// TIA Portal V18 program export: 5 tag tables, 14 data types, 1 data blocks, 8 code blocks (in call order from the OBs), 0 instance data blocks

VAR_GLOBAL   // PLC tag table "BYPASS_APERTADEIRAS"
   start AT %I1500.1 : Bool;
   remover AT %I1500.2 : Bool;
   reset AT %I1500.3 : Bool;
   MOD1_OK AT %Q1594.0 : Bool;
   MOD2_OK AT %Q1594.1 : Bool;
   RESET_MOD_1 AT %M9.1 : Bool;
   RESET_MOD_2 AT %M9.2 : Bool;
   VALIDACA0_MOD1 AT %M9.6 : Bool;
   VALIDAÇÃO_MOD2 AT %M12.0 : Bool;
   VALIDACAO_ANDON_MOD2 AT %M12.2 : Bool;
   VALIDACAO_ANDON_MOD1 AT %M12.3 : Bool;
   LEANDRO AT %M12.4 : Bool;
   BYPASS_ABST_OLEO AT %M12.6 : Bool;
   BYPASS_ABSTECIMENTO_OLEO AT %M12.7 : Bool;
   BYPASS_ESTANQ_CIL AT %M13.0 : Bool;
   BYPASS_SUP_FREIO AT %M2.1 : Bool;
   BYPASS_PY_EXCENTRICO AT %M2.2 : Bool;
   BYPASS_AP_HARPA AT %M12.5 : Bool;
   BYPASS_BUJAO AT %M13.1 : Bool;
   BYPASS_AP_BUJAO AT %M13.2 : Bool;
   BYPASS_TUBO_RPX AT %M13.3 : Bool;
   BYPASS_AP_TUBO_RPX AT %M13.4 : Bool;
   BYPASS_MOLA_HARPA AT %M13.5 : Bool;
   BYPASS_CARCACA AT %M13.6 : Bool;
   BYPASS_AP_CARCA AT %M13.7 : Bool;
   BYPASS_TALHA_DIF AT %M28.0 : Bool;
   BYPASS_SENSOR_TALHA_DIF AT %M28.1 : Bool;
   BYPASS_PYJUNTA AT %M28.2 : Bool;
   BYPASS_PY_JUNTA AT %M28.3 : Bool;
   BYPASS_CRAWFOOT AT %M28.4 : Bool;
   BYPASS_AP_CRAWFOOT AT %M28.5 : Bool;
   BYPASS_DUPLO_FUSO AT %M28.6 : Bool;
   BYPASS_AP_DUPLO_FUSO AT %M28.7 : Bool;
   BYPASS_P_ESCONDIDA AT %M29.0 : Bool;
   BYPASS_AP_PORCA_ESCON AT %M29.1 : Bool;
   BYPASS_SUP_CIL AT %M29.2 : Bool;
   BYPASS_AP_SUP_CIL AT %M29.3 : Bool;
   BYPASS_PORCA_CIL AT %M29.4 : Bool;
   BYPASS_AP_PORCA_CIL AT %M29.5 : Bool;
   BYPASS_AP_SUP_FREIO AT %M29.6 : Bool;
   BYPASS_PYEXCENTRICO AT %M29.7 : Bool;
   BYPASS_CUBO_DISC AT %M30.0 : Bool;
   BYPASS_PY_CUBO_DISC AT %M30.1 : Bool;
   BYPASS_HOLDER AT %M30.2 : Bool;
   BYPASS_AP_HOLDER AT %M30.3 : Bool;
   BYPASS_CALIPER AT %M30.4 : Bool;
   BYPASS_AP_CALPER AT %M30.5 : Bool;
   BYPASS_PYCUBO_TAMBOR AT %M30.6 : Bool;
   BYPASS_PY_CUBO_TAMBOR AT %M30.7 : Bool;
   BYPASS_HASTE_ALV AT %M31.0 : Bool;
   BYPASS_AP_HASTE_ALV AT %M31.1 : Bool;
   BYPASS_APCUBO AT %M31.2 : Bool;
   BYPASS_AP_CUBO AT %M31.3 : Bool;
   BYPASS_CRAVADOR AT %M31.4 : Bool;
   BYPASS_AP_CRAVADOR AT %M31.5 : Bool;
   BYPASS_INDICADOR AT %M31.6 : Bool;
   BYPASS_AP_INDICADOR AT %M31.7 : Bool;
   BYPASS_VALVULA AT %M32.0 : Bool;
   BYPASS_AP_VALVULA AT %M32.1 : Bool;
   BYPASS_HELGE AT %M32.2 : Bool;
   BYPASS_PY_HELGE AT %M32.3 : Bool;
   BYPASS_PORCA_TERMINAL AT %M32.4 : Bool;
   BYPASS_AP_PORCA_TERMINAL AT %M32.5 : Bool;
   BYPASS_FILTRO_OLEO AT %M32.6 : Bool;
   BYPASS_AP_FILTRO_OLEO AT %M32.7 : Bool;
   BYPASS_REDUCAO AT %M33.0 : Bool;
   BYPASS_AP_REDUCAO AT %M33.1 : Bool;
   BYPASS_FLANGE AT %M33.2 : Bool;
   BYPASS_AP_FLANGE AT %M33.3 : Bool;
   BYPASS_ESTANQ_CILINDRO AT %M33.4 : Bool;
   BYPASS_ESTANQ_CARC AT %M33.5 : Bool;
   BYPASS_ESTANQ_CARCACA AT %M33.6 : Bool;
   EMERG_CABINE_ACIONADA AT %M35.1 : Bool;
   BYPASS_VALVULA_P50 AT %M35.6 : Bool;
   BYPASS_TAMPA_CALIPER_1 AT %M36.0 : Bool;
   BYPASS_AP_VALVULA_P50 AT %M36.1 : Bool;
   TESTE_LEITOR AT %M42.4 : Bool;
   IG_CONTROL_T AT %M43.7 : Bool;
   ABORTA_P05 AT %M2.5 : Bool;
   ABORTA_JOB_P05 AT %M2.6 : Bool;
   TORQUE_ATLAS6000_P15 AT %MD48 : Real;
   PULSO_BORDA_BYPASS AT %M3.1 : Bool;
   BORDA_BYPASS_AP AT %M3.2 : Bool;
   TORQUE_DUPLO_FUSO1 AT %MD52 : Real;
   AUX_APDP AT %M3.4 : Bool;
   SIGNAL_LOST_POKA_JUNTA AT %M3.5 : Bool;
   aux_inicio_receita_pky_p30 AT %M3.7 : Bool;
   JOBOK_POKA_JUNTA_P30 AT %M4.0 : Bool;
   BYPASS_TORQUIMETRO_DIGITAL_1 AT %M4.1 : Bool;
   BYPASS_REULAGEM_ALAVANCA_1 AT %M4.5 : Bool;
   antecipa_expedicao AT %M4.6 : Bool;
   SIGINAL_LOST_PCUBO AT %M5.0 : Bool;
   pulso_teste AT %M5.7 : Bool;
   JOBDONE_ABSTECIMENTO_OLEO AT %M7.3 : Bool;
   SIGNAL_LOST_ABAST_OLEO AT %M7.4 : Bool;
   Bypass_oring_P100 AT %M7.5 : Bool;
   BYPASS_ORING_MAP_P100 AT %M8.1 : Bool;
   SIGNAL_LOST_ORING_MAP AT %M8.3 : Bool;
   InputAuxEdi AT %M8.7 : Bool;
   InputAuxEtr AT %M9.0 : Bool;
   SEM_JOB_PY_OLEO AT %M56.6 : Bool;
   JOB_PY_OLEO AT %M56.7 : Bool;
   JOBDONE_PY_GRAXA AT %M57.2 : Bool;
   Bypass_jidoka_filtro AT %M57.3 : Bool;
   BYPASS_JIDOKA_FILTRO_OLEO_P125 AT %M57.4 : Bool;
   Bypass_vaselina AT %M57.5 : Bool;
   JobOK_vaselina AT %M57.6 : Bool;
   BYpassVaselina AT %M57.7 : Bool;
   resetsinais AT %M58.0 : Bool;
   Bypass_apcilin_pneumatico AT %M58.2 : Bool;
   Bypass_apcilin_pneumaticoP105 AT %M58.3 : Bool;
END_VAR

VAR_GLOBAL   // PLC tag table "BYPASS_STATIONS"
   BYPASS_STATION_1 AT %M36.2 : Bool;
   BYPASS_POSTO_1 AT %M36.3 : Bool;
   BYPASS_STATION_5 AT %M36.4 : Bool;
   BYPASS_POSTO_5 AT %M36.5 : Bool;
   BYPASS_STATION_10 AT %M36.6 : Bool;
   BYPASS_POSTO_10 AT %M36.7 : Bool;
   BYPASS_STATION_15 AT %M37.0 : Bool;
   BYPASS_POSTO_15 AT %M37.1 : Bool;
   BYPASS_STATION_20 AT %M37.2 : Bool;
   BYPASS_POSTO_20 AT %M37.3 : Bool;
   BYPASS_STATION_30 AT %M37.4 : Bool;
   BYPASS_POSTO_30 AT %M37.5 : Bool;
   BYPASS_STATION_40 AT %M37.6 : Bool;
   BYPASS_POSTO_40 AT %M37.7 : Bool;
   BYPASS_STATION_50 AT %M38.0 : Bool;
   BYPASS_POSTO_50 AT %M38.1 : Bool;
   BYPASS_STATION_55 AT %M38.2 : Bool;
   BYPASS_POSTO_55 AT %M38.3 : Bool;
   BYPASS_STATION_60 AT %M38.4 : Bool;
   BYPASS_POSTO_60 AT %M38.5 : Bool;
   BYPASS_STATION_70 AT %M38.6 : Bool;
   BYPASS_POSTO_70 AT %M38.7 : Bool;
   BYPASS_STATION_75 AT %M39.0 : Bool;
   BYPASS_POSTO_75 AT %M39.1 : Bool;
   BYPASS_STATION_80 AT %M39.2 : Bool;
   BYPASS_POSTO_80 AT %M39.3 : Bool;
   BYPASS_STATION_90 AT %M39.4 : Bool;
   BYPASS_POSTO_90 AT %M39.5 : Bool;
   BYPASS_STATION_95 AT %M39.6 : Bool;
   BYPASS_POSTO_95 AT %M39.7 : Bool;
   BYPASS_STATION_100 AT %M40.0 : Bool;
   BYPASS_POSTO_100 AT %M40.1 : Bool;
   BYPASS_STATION_105 AT %M40.2 : Bool;
   BYPASS_POSTO_105 AT %M40.3 : Bool;
   BYPASS_STATION_110 AT %M40.4 : Bool;
   BYPASS_POSTO_110 AT %M40.5 : Bool;
   BYPASS_STATION_115 AT %M40.6 : Bool;
   BYPASS_POSTO_115 AT %M40.7 : Bool;
   BYPASS_STATION_120 AT %M41.0 : Bool;
   BYPASS_POSTO_120 AT %M41.1 : Bool;
   BYPASS_STATION_125 AT %M41.2 : Bool;
   BYPASS_POSTO_125 AT %M41.3 : Bool;
   BYPASS_STATION_130 AT %M41.4 : Bool;
   BYPASS_POSTO_130 AT %M41.5 : Bool;
   BYPASS_STATION_140 AT %M41.6 : Bool;
   BYPASS_POSTO_140 AT %M41.7 : Bool;
   BYPASS_STATION_150 AT %M42.0 : Bool;
   BYPASS_POSTO_150 AT %M42.1 : Bool;
   BYPASS_STATION_QG AT %M42.2 : Bool;
   BYPASS_POSTO_QG AT %M42.3 : Bool;
END_VAR

VAR_GLOBAL   // PLC tag table "Default tag table"
   Forced_WO AT %I1500.0 : Bool;
   Trig_Buffer_ADIC AT %I1500.4 : Bool;
   Trig_Buffer_REMOV AT %I1500.5 : Bool;
   senor_filtro_oleo AT %I1000.0 : Bool;
   LEITOR_LEN AT %IB2283 : Byte;
   LEITURA_DONE AT %I2002.4 : Bool;
   sensor_vaselina AT %I1000.4 : Bool;
   Gatilho_ap_pneumaticaP105 AT %I221.6 : Bool;
   Sensor_RX1_RBX1 AT %I201.7 : Bool;
   Sensor_RX2_RBX2 AT %I201.6 : Bool;
   Sensor_cotovelo_mangueira AT %I1050.0 : Bool;
   Sensor_cotovelo AT %I1050.2 : Bool;
   Sensor_cotovelo_AD1600 AT %I1050.4 : Bool;
   Sensor_plug AT %I1050.6 : Bool;
   Tag_1 AT %QD1302 : DWord;
   Tag_2 AT %Q400.0 : Bool;
   Tag_3 AT %QW1310 : Int;
   SINAL_AP_SEMPRE_LIGADO AT %Q4000.0 : Bool;
   Tag_4 AT %QB1100 : Byte;
   RESET_DESOUTTER_P50 AT %Q8000.0 : Bool;
   RESET_DESOUTTER_P40 AT %Q6000.0 : Bool;
   Limpa_leitor AT %Q2000.7 : Bool;
   Buzzer_P01 AT %Q3.4 : Bool;
   Led_azul_P01 AT %Q3.2 : Bool;
   Led_red_P01 AT %Q3.0 : Bool;
   Led_verde_P01 AT %Q3.1 : Bool;
   Ledverde AT %Q1000.2 : Bool;
   Ledlaranja AT %Q1000.3 : Bool;
   LedVerde_vaselina AT %Q1000.6 : Bool;
   LedAmarelo_vaselina AT %Q1000.7 : Bool;
   LED_RX1_RBX1 AT %Q200.7 : Bool;
   LED_RX2_RBX2 AT %Q200.6 : Bool;
   Buzzer_P40 AT %Q5.4 : Bool;
   Led_azulP40 AT %Q5.2 : Bool;
   Led_VermelhoP40 AT %Q5.0 : Bool;
   Led_VerdeP40 AT %Q5.1 : Bool;
   Led_cotovelo_mangueira AT %Q1050.1 : Bool;
   Led_Cotovelo AT %Q1050.3 : Bool;
   Led_cotovelo_AD1600 AT %Q1050.5 : Bool;
   Led_Plug AT %Q1050.7 : Bool;
   FirstScan AT %M1.0 : Bool;
   DiagStatusUpdate AT %M1.1 : Bool;
   AlwaysTRUE AT %M1.2 : Bool;
   AlwaysFALSE AT %M1.3 : Bool;
   Clock_Byte AT %MB0 : Byte;
   Clock_10Hz AT %M0.0 : Bool;
   Clock_5Hz AT %M0.1 : Bool;
   "Clock_2.5Hz" AT %M0.2 : Bool;
   Clock_2Hz AT %M0.3 : Bool;
   "Clock_1.25Hz" AT %M0.4 : Bool;
   Clock_1Hz AT %M0.5 : Bool;
   "Clock_0.625Hz" AT %M0.6 : Bool;
   "Clock_0.5Hz" AT %M0.7 : Bool;
   status_10 AT %M1.4 : Bool;
   status_20 AT %M1.5 : Bool;
   status_40 AT %M1.6 : Bool;
   status_50 AT %M1.7 : Bool;
   status_60 AT %M6.0 : Bool;
   status_70 AT %M6.1 : Bool;
   status_80 AT %M6.2 : Bool;
   status_90 AT %M6.3 : Bool;
   status_100 AT %M6.4 : Bool;
   status_110 AT %M6.5 : Bool;
   status_120 AT %M6.6 : Bool;
   status_130 AT %M6.7 : Bool;
   BUSY AT %M7.6 : Bool;
   CYCLE_DONE_AREA_IHM AT %M8.0 : Bool;
   MODEZONE_DONE_AREA_IHM AT %M8.2 : Bool;
   CYCLE_DONE_IT_IHM AT %M8.4 : Bool;
   BOTAO_ACIONAR_MENSAGENS AT %M8.5 : Bool;
   Quantity_ok AT %MW10 : Int;
   BYPASSLEITOR AT %M7.7 : Bool;
   Inicia_apertadeiras AT %M4.4 : Bool;
   FORÇA_RECEITA_GERAL AT %M12.1 : Bool;
   CU_PRIMEIRO_POSTO AT %MW14 : Int;
   "POPID_INICO DE_LINHA" AT %M18.0 : LInt;
   Ready_to_copy AT %M2.0 : Bool;
   BYPASS_MOD_2 AT %M2.3 : Bool;
   BYPASS_MOD_1 AT %M2.4 : Bool;
   BYPASS_GERAL_EQUIP AT %M900.1 : Bool;
   "NOVO TESTE" AT %M9.5 : Bool;
   BYPASS_GERAL AT %M33.7 : Bool;
   ESVAZIAMENTO_FALCARE AT %M34.0 : Bool;
   ESVAZIA_FALCARE AT %M34.1 : Bool;
   ESVAZIA_MAIN_LINE AT %M34.2 : Bool;
   ESVAZIAMENTO_MAIN_LINE AT %M34.3 : Bool;
   ESVAZIA_FALCARE_1 AT %M34.4 : Bool;
   ESVAZIA_MAIN_LINE_1 AT %M34.5 : Bool;
   ERRO_ESVAZIAMENTO_LINHA AT %M34.6 : Bool;
   "CABINE EM MANUAL" AT %M34.7 : Bool;
   PRODUCAO_CONCLUIDA AT %M35.0 : Bool;
   GAP_E_EIXO_PENDURADO AT %M35.2 : Bool;
   VALIDACAO_EMERG_MOD1 AT %M35.3 : Bool;
   VALIDACAO_EMERG_MOD2 AT %M35.4 : Bool;
   "SINAL_DE RESET_GAP_CABINE" AT %M35.5 : Bool;
   BYPASS_TAMPA_CALIPER AT %M35.7 : Bool;
   INDEX_LEITOR AT %MW44 : UInt;
   CARACTER AT %MW46 : Int;
   RET_VAL AT %MW200 : Int;
   BYPASS_CABINE_EM_MODO_LOCAL AT %M42.5 : Bool;
   BYPASS_CAB_MODO_LOCAL AT %M42.6 : Bool;
   ACIONA_TELA AT %M43.1 : Bool;
   ERROR_COMUNICACAO_CABINE_SEND AT %M43.2 : Bool;
   ERROR_COMUNICACAO_CABINE_RECIVE AT %M43.3 : Bool;
   BYPASS_LEITURA AT %M43.4 : Bool;
   BORDA_MODZ1 AT %M43.5 : Bool;
   BYPASS_PY_JUNTA_RX_RBX AT %M43.6 : Bool;
   bypass_sem_receita AT %M2.7 : Bool;
   provisorio AT %M3.0 : Bool;
   BYPASS_PRENSA_LEMARB AT %M3.3 : Bool;
   TOOLRUNNING_POKA_JUNTA AT %M3.6 : Bool;
   BYPASS_TORQUIMETRO_DIGITAL AT %M4.2 : Bool;
   BYPASS_REULAGEM_ALAVANCA AT %M4.3 : Bool;
   ATIVA_FOR AT %M4.7 : Bool;
   PULSO_BY_P110 AT %M5.1 : Bool;
   set_modezone_done AT %M5.2 : Bool;
   giro_cabine AT %M5.3 : Bool;
   cabine_rodou AT %M5.4 : Bool;
   reset_md1 AT %M5.5 : Bool;
   reset_md2 AT %M5.6 : Bool;
   aux_gap AT %M7.0 : Bool;
   guarda_gap AT %M7.1 : Bool;
   chamada_forcada AT %MW16 : Int;
   Cabin_line_reference AT %M7.2 : Bool;
   SIGNAL_LOST_HELGE_2 AT %M8.6 : Bool;
   Habilita_matrix_P01 AT %M9.3 : Bool;
   Habilita_matrix_P05 AT %M9.4 : Bool;
   Habilita_matrix_P10 AT %M9.7 : Bool;
   Habilita_matrix_P15 AT %M26.0 : Bool;
   Habilita_matrix_P20 AT %M26.1 : Bool;
   Habilita_matrix_P30 AT %M26.2 : Bool;
   Habilita_matrix_P40 AT %M26.3 : Bool;
   Habilita_matrix_P50 AT %M26.4 : Bool;
   Habilita_matrix_P55 AT %M26.5 : Bool;
   Habilita_matrix_P60 AT %M26.6 : Bool;
   Habilita_matrix_P70 AT %M26.7 : Bool;
   Habilita_matrix_P75 AT %M27.0 : Bool;
   Habilita_matrix_P80 AT %M27.1 : Bool;
   Habilita_matrix_P90 AT %M27.2 : Bool;
   Habilita_matrix_P95 AT %M27.3 : Bool;
   Habilita_matrix_P100 AT %M27.4 : Bool;
   Habilita_matrix_P105 AT %M27.5 : Bool;
   Habilita_matrix_P110 AT %M27.6 : Bool;
   Habilita_matrix_P115 AT %M27.7 : Bool;
   Habilita_matrix_P120 AT %M42.7 : Bool;
   Habilita_matrix_P125 AT %M43.0 : Bool;
   Habilita_matrix_P130 AT %M56.0 : Bool;
   Habilita_matrix_P140 AT %M56.1 : Bool;
   Habilita_matrix_P150 AT %M56.2 : Bool;
   Habilita_matrix_QG AT %M56.3 : Bool;
   Bypass_graxa AT %M56.4 : Bool;
   Bypass_graxa_expedicao AT %M56.5 : Bool;
   JOBOK_PY_OLEO AT %M57.0 : Bool;
   antecipa_expedicao_1 AT %M57.1 : Bool;
   bahia AT %M58.1 : Bool;
   Count_gatilho AT %MW60 : Int;
END_VAR
VAR_GLOBAL CONSTANT   // user constants
   Config_OPC : Int := 17;
   maxConnectionsOPCUA : Int := 5;
END_VAR

VAR_GLOBAL   // PLC tag table "LEITOR_VIVERK"
   Readcomplete AT %I2000.1 : Bool;
   ResultData0 AT %IB2284 : Byte;
   ResultData1 AT %IB2285 : Byte;
   ResultData2 AT %IB2286 : Byte;
   ResultData3 AT %IB2287 : Byte;
   ResultData4 AT %IB2288 : Byte;
   ResultData5 AT %IB2289 : Byte;
   ResultData6 AT %IB2290 : Byte;
   ResultData7 AT %IB2291 : Byte;
   ResultData8 AT %IB2292 : Byte;
   ResultData9 AT %IB2293 : Byte;
   ResultData10 AT %IB2294 : Byte;
   ResultData11 AT %IB2295 : Byte;
   ResultData12 AT %IB2296 : Byte;
   Tag_5 AT %IB2000 : Byte;
   Tag_6 AT %IB2001 : Byte;
   Tag_7 AT %IB2002 : Byte;
   Tag_8 AT %IB2003 : Byte;
   Tag_9 AT %IB2004 : Byte;
   Tag_10 AT %IB2005 : Byte;
   Tag_11 AT %IB2006 : Byte;
   Tag_12 AT %IB2007 : Byte;
   Tag_13 AT %IB2008 : Byte;
   Tag_14 AT %IB2009 : Byte;
   Tag_15 AT %IB2010 : Byte;
   Tag_16 AT %IB2011 : Byte;
   Tag_17 AT %IB2012 : Byte;
   Tag_18 AT %IB2013 : Byte;
END_VAR

VAR_GLOBAL   // PLC tag table "Setup"
   Tag_19 AT %I0.0 : Bool;
END_VAR
VAR_GLOBAL CONSTANT   // user constants
   ModeZone_Setup_Const : Int := 12;
   Station_Setup_Const : Int := 20;
   Position_Setup_Const : Int := 1;
   Equipment_Setup_Const : Int := 10;
   ThisProcess : Int := 1;
   ThisWorkshop : Int := 1;
   Connection_Setup_Const : Int := 30;
   ContractID_Setup_Const : Int := 24;
   ITConnectionName : String := 'PLC_AREA_01';
   Parameter_Setup_Const : Int := 20;
   WorkPlace_Setup_Const : Int := 16;
   Total_User_Const : Int := 200;
   User_Roles_Const : Int := 100;
   ProductionSequenceList_Setup_Const : Int := 30;   // Quantidade de produtos que podemos ter por posto
   listTypeReason_Const : Int := 200;
   ITConnectionID : Word := W#16#101;
   Signal_Setup_Const : Int := 8;
   ShiftList_Setup_Const : Int := 3;
   Quantidade_task : Int := 10;
   Tamanho_POPID : Int := 7;
   nProcess : Int := 1;
   Quantidade_Paradas_Matriz : Int := 2;
END_VAR

TYPE "Comm"
   STRUCT
      Connection_ID : Word;
      R_ID : CONN_R_ID;
      REQ : Bool;
      Len : Word;
      Result : Struct
         DONE : Bool;
         ERROR : Bool;
         STATUS : Word;
      END_STRUCT;
      Diagnostic : Struct
         countDone : Int;
         countError : Int;
         memStatus : Word;
      END_STRUCT;
   END_STRUCT;
END_TYPE

TYPE "Config_SEND_RCV"
   STRUCT
      modezone { S7_SetPoint := 'True'} : Array[1.."ModeZone_Setup_Const"] of "Comm";
   END_STRUCT;
END_TYPE

TYPE "InterlockEmergMdz_in"
   STRUCT
      StationInterlock_APLC_Input : Array[1.."Station_Setup_Const"] of Struct
         Emergencial_Interlock_APLC_Input : Bool;
      END_STRUCT;
   END_STRUCT;
END_TYPE

TYPE "InterlockMdz_in"
   STRUCT
      StationInterlock_APLC_Input : Array[1.."Station_Setup_Const"] of Struct
         PositionInterlock_APLC_Input : Array[1.."Position_Setup_Const"] of Struct
            LoginInterlock_APLC : Bool;
            EquipmentInterlock_APLC_Input : Array[1.."Equipment_Setup_Const"] of Struct
               SignalInterlock_APLC_Input : Array[1.."Signal_Setup_Const"] of Bool;
            END_STRUCT;
         END_STRUCT;
      END_STRUCT;
   END_STRUCT;
END_TYPE

TYPE "Modezone_Gap"
   STRUCT
      GapActive : Bool;
   END_STRUCT;
END_TYPE

TYPE "Process_Gap"
   STRUCT
      ProcessGapActive : Bool;
      ModezoneGap { S7_SetPoint := 'True'} : Array[1.."ModeZone_Setup_Const"] of "Modezone_Gap";
   END_STRUCT;
END_TYPE

TYPE "TaktModeZone_Input"
   STRUCT
      ModeZone_Done : Bool;
   END_STRUCT;
END_TYPE

TYPE "TargetProductionMdz_in"
   STRUCT
      KPI_Informations : Struct
         Full_AvailabilityShift : Array[1.."ShiftList_Setup_Const"] of Time;
         Full_AvailabilityDay : Time := T#9H_15M;
         Net_AvailabilityShift : Array[1.."ShiftList_Setup_Const"] of Time;
         Net_AvailabilityDay : Time := T#9H_15M;
         Total_StopPlannedShift : Array[1.."ShiftList_Setup_Const"] of Time;
         Total_StopPlannedDay : Time := T#0MS;
         StopPlanned_Executed_Shift : Array[1.."ShiftList_Setup_Const"] of Time;
         StopPlanned_Executed_Day : Time := T#2H_45M;
         NextStopPlanned : Date_And_Time := DT#2000-01-10-00:00:00;
         NextStopPlanned_Index : Int := 11;
         RemaningTimeToStopPlanned : Time := T#8D_15H_45M_48S_109MS;
         NextStopPlannedInRealTime : Time := T#8H_14M_11S_891MS;
         RemaningCycleToStoPplanned : DInt := 2_139_095_040;
         Total_StopTimeShift : Array[1.."ShiftList_Setup_Const"] of Time;
         Total_StopTimeDay : Time := T#-1H_41M_28S;
         GoalOfShift : Array[1.."ShiftList_Setup_Const"] of Int;
         GoalOfDay : Int := 199;
         TaktStandardByShift : Array[1.."ShiftList_Setup_Const"] of Time;
      END_STRUCT;
      KPI_Results : Struct
         Production_Status : Int := 0;
         MaxProductionCapacity_Shift : Array[1.."ShiftList_Setup_Const"] of Int;
         MaxProductionCapacity_Day : Int := 246;
         TimeToProductionDone_Shift : Array[1.."ShiftList_Setup_Const"] of Time;
         TimeToProductionDone_Day : Time := T#0MS;
      END_STRUCT;
   END_STRUCT;
   // KPI_Informations.Full_AvailabilityShift[1] := T#9H_15M;
   // KPI_Informations.Full_AvailabilityShift[2..3] := T#0MS;
   // KPI_Informations.Net_AvailabilityShift[1] := T#9H_15M;
   // KPI_Informations.Net_AvailabilityShift[2..3] := T#0MS;
   // KPI_Informations.Total_StopPlannedShift[1..3] := T#0MS;
   // KPI_Informations.StopPlanned_Executed_Shift[1] := T#1H_35M;
   // KPI_Informations.StopPlanned_Executed_Shift[2] := T#1H_10M;
   // KPI_Informations.StopPlanned_Executed_Shift[3] := T#0MS;
   // KPI_Informations.Total_StopTimeShift[1] := T#-1H_11M_58S;
   // KPI_Informations.Total_StopTimeShift[2] := T#-29M_30S;
   // KPI_Informations.Total_StopTimeShift[3] := T#0MS;
   // KPI_Informations.GoalOfShift[1] := 164;
   // KPI_Informations.GoalOfShift[2] := 35;
   // KPI_Informations.GoalOfShift[3] := 0;
   // KPI_Informations.TaktStandardByShift[1] := T#2M_15S;
   // KPI_Informations.TaktStandardByShift[2] := T#10M;
   // KPI_Informations.TaktStandardByShift[3] := T#0MS;
   // KPI_Results.MaxProductionCapacity_Shift[1] := 246;
   // KPI_Results.MaxProductionCapacity_Shift[2..3] := 0;
   // KPI_Results.TimeToProductionDone_Shift[1..3] := T#0MS;
END_TYPE

TYPE "UDT_DadosEquipScala"
   STRUCT
      Bool0 : Bool;
      Bool1 : Bool;
      Bool2 : Bool;
      Bool3 : Bool;
      Bool4 : Bool;
      Bool5 : Bool;
      Bool6 : Bool;
      Bool7 : Bool;
      Bool8 : Bool;
      Bool9 : Bool;
      Bool10 : Bool;
      Bool11 : Bool;
      Bool12 : Bool;
      Bool13 : Bool;
      Bool14 : Bool;
      Bool15 : Bool;
   END_STRUCT;
END_TYPE

TYPE "UDT_EquipamentoScala"
   STRUCT
      Equipamento : Array[1..18] of "UDT_DadosEquipScala";
   END_STRUCT;
END_TYPE

TYPE "Udt_DataAGVStation"
   STRUCT
      Station { S7_SetPoint := 'True'} : Array[1..20] of "Udt_Data_AGVToScala";
   END_STRUCT;
END_TYPE

TYPE "Udt_Data_AGVToScala"
   STRUCT
      POPID : String[10];   // POPID
      CU : String[10];   // CU
      AGVNumber : Int;   // Número AGV
      ProductOK : Bool;   // Produto recebido OK
      ProductNOK : Bool;   // Falha produto recebido Scala
      AGVRedCard : Bool;   // AGV com trabalho
      Spare4 : Bool;   // Reserva
      Spare5 : Bool;   // Reserva
      Spare6 : Bool;   // Reserva
      Spare7 : Bool;   // Reserva
      Spare8 : Bool;   // Reserva
      Spare9 : Bool;   // Reserva
      Spare10 : Bool;   // Reserva
      Spare11 : Bool;   // Reserva
      Spare12 : Bool;   // Reserva
      Spare13 : Bool;   // Reserva
      Spare14 : Bool;   // Reserva
      Spare15 : Bool;   // Reserva
      Spare16 : Bool;   // Reserva
   END_STRUCT;
END_TYPE

TYPE "UserValidationMdz_in"
   STRUCT
      Station : Array[1.."Station_Setup_Const"] of Struct
         UserMaster_ID : DInt;
         Position_ID_Validation : Int;
         LogIn : Bool;
         Position : Array[1.."Position_Setup_Const"] of Struct
            User_ID : DInt;
            BadgeNumber : LInt;
            LogIn : Bool;
            LogOut : Bool;
            ByPass : Bool;
         END_STRUCT;
      END_STRUCT;
   END_STRUCT;
   // Station[1..20].UserMaster_ID := 0;
   // Station[1..20].Position_ID_Validation := 0;
   // Station[1..20].LogIn := FALSE;
   // Station[1].Position[1].User_ID := 0;
   // Station[2].Position[1].User_ID := 0;
   // Station[3].Position[1].User_ID := 0;
   // Station[4].Position[1].User_ID := 0;
   // Station[5].Position[1].User_ID := 0;
   // Station[6].Position[1].User_ID := 0;
   // Station[7].Position[1].User_ID := 0;
   // Station[8].Position[1].User_ID := 0;
   // Station[9].Position[1].User_ID := 0;
   // Station[10].Position[1].User_ID := 0;
   // Station[11].Position[1].User_ID := 0;
   // Station[12].Position[1].User_ID := 0;
   // Station[13].Position[1].User_ID := 0;
   // Station[14].Position[1].User_ID := 0;
   // Station[15].Position[1].User_ID := 0;
   // Station[16].Position[1].User_ID := 0;
   // Station[17].Position[1].User_ID := 0;
   // Station[18].Position[1].User_ID := 0;
   // Station[19].Position[1].User_ID := 0;
   // Station[20].Position[1].User_ID := 0;
   // Station[1].Position[1].BadgeNumber := 0;
   // Station[2].Position[1].BadgeNumber := 0;
   // Station[3].Position[1].BadgeNumber := 0;
   // Station[4].Position[1].BadgeNumber := 0;
   // Station[5].Position[1].BadgeNumber := 0;
   // Station[6].Position[1].BadgeNumber := 0;
   // Station[7].Position[1].BadgeNumber := 0;
   // Station[8].Position[1].BadgeNumber := 0;
   // Station[9].Position[1].BadgeNumber := 0;
   // Station[10].Position[1].BadgeNumber := 0;
   // Station[11].Position[1].BadgeNumber := 0;
   // Station[12].Position[1].BadgeNumber := 0;
   // Station[13].Position[1].BadgeNumber := 0;
   // Station[14].Position[1].BadgeNumber := 0;
   // Station[15].Position[1].BadgeNumber := 0;
   // Station[16].Position[1].BadgeNumber := 0;
   // Station[17].Position[1].BadgeNumber := 0;
   // Station[18].Position[1].BadgeNumber := 0;
   // Station[19].Position[1].BadgeNumber := 0;
   // Station[20].Position[1].BadgeNumber := 0;
   // Station[1].Position[1].LogIn := FALSE;
   // Station[2].Position[1].LogIn := FALSE;
   // Station[3].Position[1].LogIn := FALSE;
   // Station[4].Position[1].LogIn := FALSE;
   // Station[5].Position[1].LogIn := FALSE;
   // Station[6].Position[1].LogIn := FALSE;
   // Station[7].Position[1].LogIn := FALSE;
   // Station[8].Position[1].LogIn := FALSE;
   // Station[9].Position[1].LogIn := FALSE;
   // Station[10].Position[1].LogIn := FALSE;
   // Station[11].Position[1].LogIn := FALSE;
   // Station[12].Position[1].LogIn := FALSE;
   // Station[13].Position[1].LogIn := FALSE;
   // Station[14].Position[1].LogIn := FALSE;
   // Station[15].Position[1].LogIn := FALSE;
   // Station[16].Position[1].LogIn := FALSE;
   // Station[17].Position[1].LogIn := FALSE;
   // Station[18].Position[1].LogIn := FALSE;
   // Station[19].Position[1].LogIn := FALSE;
   // Station[20].Position[1].LogIn := FALSE;
   // Station[1].Position[1].LogOut := TRUE;
   // Station[2].Position[1].LogOut := TRUE;
   // Station[3].Position[1].LogOut := TRUE;
   // Station[4].Position[1].LogOut := TRUE;
   // Station[5].Position[1].LogOut := TRUE;
   // Station[6].Position[1].LogOut := TRUE;
   // Station[7].Position[1].LogOut := TRUE;
   // Station[8].Position[1].LogOut := TRUE;
   // Station[9].Position[1].LogOut := TRUE;
   // Station[10].Position[1].LogOut := TRUE;
   // Station[11].Position[1].LogOut := TRUE;
   // Station[12].Position[1].LogOut := TRUE;
   // Station[13].Position[1].LogOut := TRUE;
   // Station[14].Position[1].LogOut := TRUE;
   // Station[15].Position[1].LogOut := TRUE;
   // Station[16].Position[1].LogOut := TRUE;
   // Station[17].Position[1].LogOut := TRUE;
   // Station[18].Position[1].LogOut := TRUE;
   // Station[19].Position[1].LogOut := TRUE;
   // Station[20].Position[1].LogOut := TRUE;
   // Station[1].Position[1].ByPass := FALSE;
   // Station[2].Position[1].ByPass := FALSE;
   // Station[3].Position[1].ByPass := FALSE;
   // Station[4].Position[1].ByPass := FALSE;
   // Station[5].Position[1].ByPass := FALSE;
   // Station[6].Position[1].ByPass := FALSE;
   // Station[7].Position[1].ByPass := FALSE;
   // Station[8].Position[1].ByPass := FALSE;
   // Station[9].Position[1].ByPass := FALSE;
   // Station[10].Position[1].ByPass := FALSE;
   // Station[11].Position[1].ByPass := FALSE;
   // Station[12].Position[1].ByPass := FALSE;
   // Station[13].Position[1].ByPass := FALSE;
   // Station[14].Position[1].ByPass := FALSE;
   // Station[15].Position[1].ByPass := FALSE;
   // Station[16].Position[1].ByPass := FALSE;
   // Station[17].Position[1].ByPass := FALSE;
   // Station[18].Position[1].ByPass := FALSE;
   // Station[19].Position[1].ByPass := FALSE;
   // Station[20].Position[1].ByPass := FALSE;
END_TYPE

TYPE "UserValidationMdz_out"
   STRUCT
      Station : Array[1.."Station_Setup_Const"] of Struct
         Position : Array[1.."Position_Setup_Const"] of Struct
            User_ID : DInt;
            User_SSB : String[8];
            UserName : String[37];
            MsgLogin : String[40];
            AuthorizedByUserMaster_ID : DInt;
            Authentication : Bool;
         END_STRUCT;
      END_STRUCT;
   END_STRUCT;
   // Station[1].Position[1].User_ID := 0;
   // Station[2].Position[1].User_ID := 0;
   // Station[3].Position[1].User_ID := 0;
   // Station[4].Position[1].User_ID := 0;
   // Station[5].Position[1].User_ID := 0;
   // Station[6].Position[1].User_ID := 0;
   // Station[7].Position[1].User_ID := 0;
   // Station[8].Position[1].User_ID := 0;
   // Station[9].Position[1].User_ID := 0;
   // Station[10].Position[1].User_ID := 0;
   // Station[11].Position[1].User_ID := 0;
   // Station[12].Position[1].User_ID := 0;
   // Station[13].Position[1].User_ID := 0;
   // Station[14].Position[1].User_ID := 0;
   // Station[15].Position[1].User_ID := 0;
   // Station[16].Position[1].User_ID := 0;
   // Station[17].Position[1].User_ID := 0;
   // Station[18].Position[1].User_ID := 0;
   // Station[19].Position[1].User_ID := 0;
   // Station[20].Position[1].User_ID := 0;
   // Station[1].Position[1].User_SSB := '';
   // Station[2].Position[1].User_SSB := '';
   // Station[3].Position[1].User_SSB := '';
   // Station[4].Position[1].User_SSB := '';
   // Station[5].Position[1].User_SSB := '';
   // Station[6].Position[1].User_SSB := '';
   // Station[7].Position[1].User_SSB := '';
   // Station[8].Position[1].User_SSB := '';
   // Station[9].Position[1].User_SSB := '';
   // Station[10].Position[1].User_SSB := '';
   // Station[11].Position[1].User_SSB := '';
   // Station[12].Position[1].User_SSB := '';
   // Station[13].Position[1].User_SSB := '';
   // Station[14].Position[1].User_SSB := '';
   // Station[15].Position[1].User_SSB := '';
   // Station[16].Position[1].User_SSB := '';
   // Station[17].Position[1].User_SSB := '';
   // Station[18].Position[1].User_SSB := '';
   // Station[19].Position[1].User_SSB := '';
   // Station[20].Position[1].User_SSB := '';
   // Station[1].Position[1].UserName := '';
   // Station[2].Position[1].UserName := '';
   // Station[3].Position[1].UserName := '';
   // Station[4].Position[1].UserName := '';
   // Station[5].Position[1].UserName := '';
   // Station[6].Position[1].UserName := '';
   // Station[7].Position[1].UserName := '';
   // Station[8].Position[1].UserName := '';
   // Station[9].Position[1].UserName := '';
   // Station[10].Position[1].UserName := '';
   // Station[11].Position[1].UserName := '';
   // Station[12].Position[1].UserName := '';
   // Station[13].Position[1].UserName := '';
   // Station[14].Position[1].UserName := '';
   // Station[15].Position[1].UserName := '';
   // Station[16].Position[1].UserName := '';
   // Station[17].Position[1].UserName := '';
   // Station[18].Position[1].UserName := '';
   // Station[19].Position[1].UserName := '';
   // Station[20].Position[1].UserName := '';
   // Station[1].Position[1].MsgLogin := 'POSTO: 1 NAO POSSUI USUARIO CADASTRADO';
   // Station[2].Position[1].MsgLogin := 'POSTO: 1 NAO POSSUI USUARIO CADASTRADO';
   // Station[3].Position[1].MsgLogin := 'POSTO: 1 NAO POSSUI USUARIO CADASTRADO';
   // Station[4].Position[1].MsgLogin := 'POSTO: 1 NAO POSSUI USUARIO CADASTRADO';
   // Station[5].Position[1].MsgLogin := 'POSTO: 1 NAO POSSUI USUARIO CADASTRADO';
   // Station[6].Position[1].MsgLogin := 'POSTO: 1 NAO POSSUI USUARIO CADASTRADO';
   // Station[7].Position[1].MsgLogin := 'POSTO: 1 NAO POSSUI USUARIO CADASTRADO';
   // Station[8].Position[1].MsgLogin := 'POSTO: 1 NAO POSSUI USUARIO CADASTRADO';
   // Station[9].Position[1].MsgLogin := 'POSTO: 1 NAO POSSUI USUARIO CADASTRADO';
   // Station[10].Position[1].MsgLogin := 'POSTO: 1 NAO POSSUI USUARIO CADASTRADO';
   // Station[11].Position[1].MsgLogin := 'POSTO: 1 NAO POSSUI USUARIO CADASTRADO';
   // Station[12].Position[1].MsgLogin := 'POSTO: 1 NAO POSSUI USUARIO CADASTRADO';
   // Station[13].Position[1].MsgLogin := 'POSTO: 1 NAO POSSUI USUARIO CADASTRADO';
   // Station[14].Position[1].MsgLogin := 'POSTO: 1 NAO POSSUI USUARIO CADASTRADO';
   // Station[15].Position[1].MsgLogin := 'POSTO: 1 NAO POSSUI USUARIO CADASTRADO';
   // Station[16].Position[1].MsgLogin := 'POSTO: 1 NAO POSSUI USUARIO CADASTRADO';
   // Station[17].Position[1].MsgLogin := 'POSTO: 1 NAO POSSUI USUARIO CADASTRADO';
   // Station[18].Position[1].MsgLogin := 'POSTO: 1 NAO POSSUI USUARIO CADASTRADO';
   // Station[19].Position[1].MsgLogin := 'POSTO: 1 NAO POSSUI USUARIO CADASTRADO';
   // Station[20].Position[1].MsgLogin := 'POSTO: 1 NAO POSSUI USUARIO CADASTRADO';
   // Station[1].Position[1].AuthorizedByUserMaster_ID := 0;
   // Station[2].Position[1].AuthorizedByUserMaster_ID := 0;
   // Station[3].Position[1].AuthorizedByUserMaster_ID := 0;
   // Station[4].Position[1].AuthorizedByUserMaster_ID := 0;
   // Station[5].Position[1].AuthorizedByUserMaster_ID := 0;
   // Station[6].Position[1].AuthorizedByUserMaster_ID := 0;
   // Station[7].Position[1].AuthorizedByUserMaster_ID := 0;
   // Station[8].Position[1].AuthorizedByUserMaster_ID := 0;
   // Station[9].Position[1].AuthorizedByUserMaster_ID := 0;
   // Station[10].Position[1].AuthorizedByUserMaster_ID := 0;
   // Station[11].Position[1].AuthorizedByUserMaster_ID := 0;
   // Station[12].Position[1].AuthorizedByUserMaster_ID := 0;
   // Station[13].Position[1].AuthorizedByUserMaster_ID := 0;
   // Station[14].Position[1].AuthorizedByUserMaster_ID := 0;
   // Station[15].Position[1].AuthorizedByUserMaster_ID := 0;
   // Station[16].Position[1].AuthorizedByUserMaster_ID := 0;
   // Station[17].Position[1].AuthorizedByUserMaster_ID := 0;
   // Station[18].Position[1].AuthorizedByUserMaster_ID := 0;
   // Station[19].Position[1].AuthorizedByUserMaster_ID := 0;
   // Station[20].Position[1].AuthorizedByUserMaster_ID := 0;
   // Station[1].Position[1].Authentication := FALSE;
   // Station[2].Position[1].Authentication := FALSE;
   // Station[3].Position[1].Authentication := FALSE;
   // Station[4].Position[1].Authentication := FALSE;
   // Station[5].Position[1].Authentication := FALSE;
   // Station[6].Position[1].Authentication := FALSE;
   // Station[7].Position[1].Authentication := FALSE;
   // Station[8].Position[1].Authentication := FALSE;
   // Station[9].Position[1].Authentication := FALSE;
   // Station[10].Position[1].Authentication := FALSE;
   // Station[11].Position[1].Authentication := FALSE;
   // Station[12].Position[1].Authentication := FALSE;
   // Station[13].Position[1].Authentication := FALSE;
   // Station[14].Position[1].Authentication := FALSE;
   // Station[15].Position[1].Authentication := FALSE;
   // Station[16].Position[1].Authentication := FALSE;
   // Station[17].Position[1].Authentication := FALSE;
   // Station[18].Position[1].Authentication := FALSE;
   // Station[19].Position[1].Authentication := FALSE;
   // Station[20].Position[1].Authentication := FALSE;
END_TYPE

DATA_BLOCK "VERIFICA INTERLOCK"   // DB200
{ S7_Optimized_Access := 'TRUE' }
// stored: MemoryReserve 100
   VAR
      INTERLOCK : Array[0..10] of Struct
         STATION : Int;
         EQUIPAMENTO : Int;
         SINAL : Int;
      END_STRUCT;
      "ATIVA FOR" : Bool;
      modezone : Int;
   END_VAR
BEGIN
END_DATA_BLOCK

ORGANIZATION_BLOCK "OB1 Main"   // OB1, LAD, ProgramCycle
TITLE = "Main Program Sweep (Cycle)"
{ S7_Optimized_Access := 'TRUE' }
// stored: SetENOAutomatically false
   VAR_INPUT
      Initial_Call : Bool;   // Initial call of this OB
      Remanence : Bool;   // =True, if remanent data are available
   END_VAR
   VAR_TEMP
      ADR : UDInt;
      LEN : UInt;
      "RETURN" : Int;
      ERROR : Bool;
      STATUS : Word;
      DONE : Bool;
      POPID : String;
      CU : Int;
      Quantidade_erro : Int;
      DONE_MAIN_LINE_PUT : Bool;
      ERROR_MAIN_LINE_PUT : Bool;
      DONE_MAIN_LINE_GET : Bool;
      ERROR_MAIN_LINE_GET : Bool;
      DONE_FALCARE_PUT : Bool;
      ERROR_FALCARE_PUT : Bool;
      DONE_FALCARE_GET : Bool;
      ERROR_FALCARE_GET : Bool;
      DONE_GIRADOR_PUT : Bool;
      ERROR_GIRADOR_PUT : Bool;
      DONE_GIRADOR_GET : Bool;
      ERROR_GIRADOR_GET : Bool;
      DONE_ABSTECIMENTO_OLEO_PUT : Bool;
      ERRO_ABASTECIMENTO_OLEO_PUT : Bool;
      DONE_ABSTECIMENTO_OLEO_GET : Bool;
      ERRO_ABSTECIMENTO_OLEO_GET : Bool;
      ERROR_ALARMS_IHM_FALCARE_GET : Bool;
      DONE_ALARMS_IHM_FALCARE_GET : Bool;
      AUX_BSEND_LEMARB : Word;
      AUX_RECIVE_LEMARB : Word;
   END_VAR
BEGIN

REGION Network 1: Set Id Connection automatic
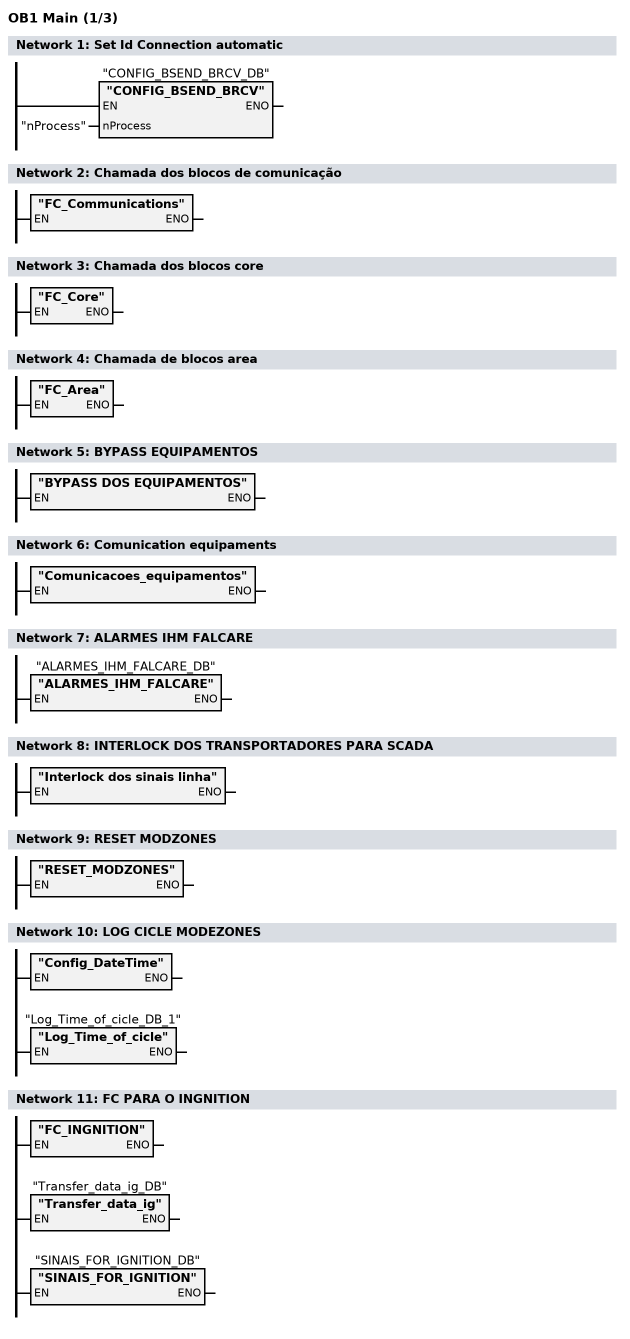
   RUNG wire#powerrail
      "CONFIG_BSEND_BRCV_DB"(nProcess := "nProcess")
   END_RUNG
   // the same network as SCL:
   "CONFIG_BSEND_BRCV_DB"(nProcess := "nProcess");   // "CONFIG_BSEND_BRCV"
END_REGION

REGION Network 2: Chamada dos blocos de comunicação
   RUNG wire#powerrail
      "FC_Communications"()
   END_RUNG
   // the same network as SCL:
   "FC_Communications"();
END_REGION

REGION Network 3: Chamada dos blocos core
   RUNG wire#powerrail
      "FC_Core"()
   END_RUNG
   // the same network as SCL:
   "FC_Core"();
END_REGION

REGION Network 4: Chamada de blocos area
   RUNG wire#powerrail
      "FC_Area"()
   END_RUNG
   // the same network as SCL:
   "FC_Area"();
END_REGION

REGION Network 5: BYPASS EQUIPAMENTOS
   RUNG wire#powerrail
      "BYPASS DOS EQUIPAMENTOS"()
   END_RUNG
   // the same network as SCL:
   "BYPASS DOS EQUIPAMENTOS"();
END_REGION

REGION Network 6: Comunication equipaments
   RUNG wire#powerrail
      "Comunicacoes_equipamentos"()
   END_RUNG
   // the same network as SCL:
   "Comunicacoes_equipamentos"();
END_REGION

REGION Network 7: ALARMES IHM FALCARE
   RUNG wire#powerrail
      "ALARMES_IHM_FALCARE_DB"()
   END_RUNG
   // the same network as SCL:
   "ALARMES_IHM_FALCARE_DB"();   // "ALARMES_IHM_FALCARE"
END_REGION

REGION Network 8: INTERLOCK DOS TRANSPORTADORES PARA SCADA
   RUNG wire#powerrail
      "Interlock dos sinais linha"()
   END_RUNG
   // the same network as SCL:
   "Interlock dos sinais linha"();
END_REGION

REGION Network 9: RESET MODZONES
   RUNG wire#powerrail
      "RESET_MODZONES"()
   END_RUNG
   // the same network as SCL:
   "RESET_MODZONES"();
END_REGION

REGION Network 10: LOG CICLE MODEZONES
   RUNG wire#powerrail
      "Config_DateTime"()
   END_RUNG
   RUNG wire#powerrail
      "Log_Time_of_cicle_DB_1"()
   END_RUNG
   // the same network as SCL:
   "Config_DateTime"();
   "Log_Time_of_cicle_DB_1"();   // "Log_Time_of_cicle"
END_REGION

REGION Network 11: FC PARA O INGNITION
   RUNG wire#powerrail
      "FC_INGNITION"()
   END_RUNG
   RUNG wire#powerrail
      "Transfer_data_ig_DB"()
   END_RUNG
   RUNG wire#powerrail
      "SINAIS_FOR_IGNITION_DB"()
   END_RUNG
   // the same network as SCL:
   "FC_INGNITION"();
   "Transfer_data_ig_DB"();   // "Transfer_data_ig"
   "SINAIS_FOR_IGNITION_DB"();   // "SINAIS_FOR_IGNITION"
END_REGION

REGION Network 12: TESTE DE VALIDAÇÃO MODEZONES
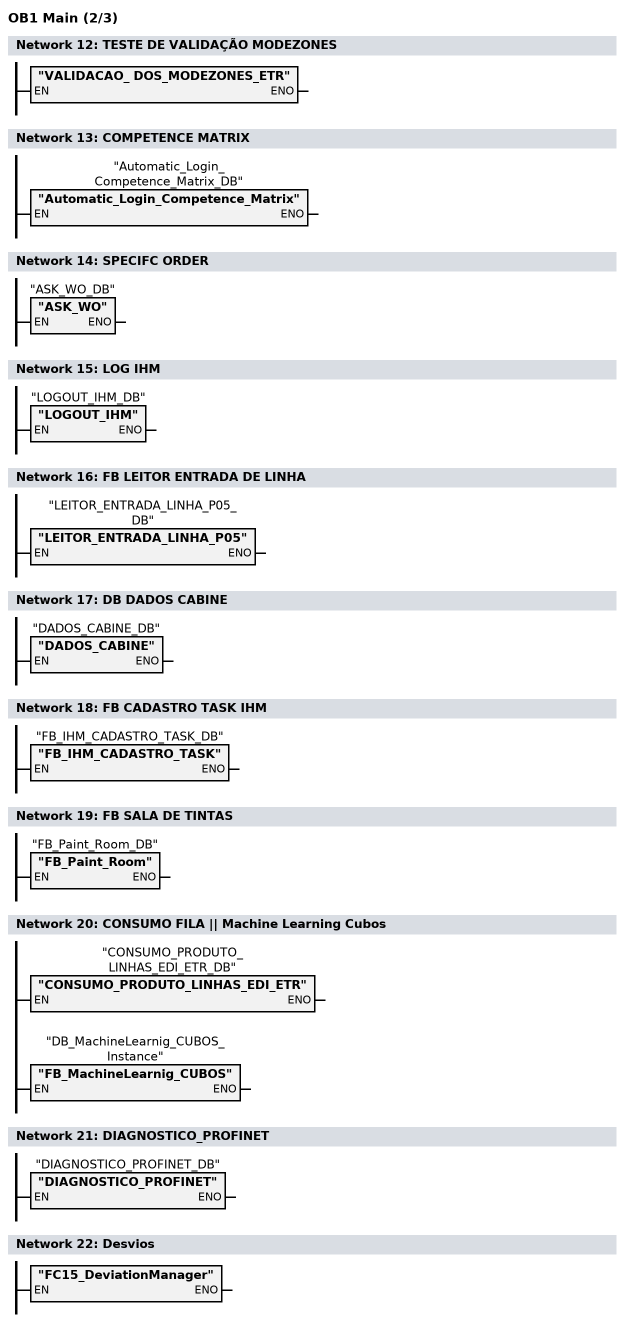
   RUNG wire#powerrail
      "VALIDACAO_ DOS_MODEZONES_ETR"()
   END_RUNG
   // the same network as SCL:
   "VALIDACAO_ DOS_MODEZONES_ETR"();
END_REGION

REGION Network 13: COMPETENCE MATRIX
   RUNG wire#powerrail
      "Automatic_Login_Competence_Matrix_DB"()
   END_RUNG
   // the same network as SCL:
   "Automatic_Login_Competence_Matrix_DB"();   // "Automatic_Login_Competence_Matrix"
END_REGION

REGION Network 14: SPECIFC ORDER
   RUNG wire#powerrail
      "ASK_WO_DB"()
   END_RUNG
   // the same network as SCL:
   "ASK_WO_DB"();   // "ASK_WO"
END_REGION

REGION Network 15: LOG IHM
   RUNG wire#powerrail
      "LOGOUT_IHM_DB"()
   END_RUNG
   // the same network as SCL:
   "LOGOUT_IHM_DB"();   // "LOGOUT_IHM"
END_REGION

REGION Network 16: FB LEITOR ENTRADA DE LINHA
   RUNG wire#powerrail
      "LEITOR_ENTRADA_LINHA_P05_DB"()
   END_RUNG
   // the same network as SCL:
   "LEITOR_ENTRADA_LINHA_P05_DB"();   // "LEITOR_ENTRADA_LINHA_P05"
END_REGION

REGION Network 17: DB DADOS CABINE
   RUNG wire#powerrail
      "DADOS_CABINE_DB"()
   END_RUNG
   // the same network as SCL:
   "DADOS_CABINE_DB"();   // "DADOS_CABINE"
END_REGION

REGION Network 18: FB CADASTRO TASK IHM
   RUNG wire#powerrail
      "FB_IHM_CADASTRO_TASK_DB"()
   END_RUNG
   // the same network as SCL:
   "FB_IHM_CADASTRO_TASK_DB"();   // "FB_IHM_CADASTRO_TASK"
END_REGION

REGION Network 19: FB SALA DE TINTAS
   RUNG wire#powerrail
      "FB_Paint_Room_DB"()
   END_RUNG
   // the same network as SCL:
   "FB_Paint_Room_DB"();   // "FB_Paint_Room"
END_REGION

REGION Network 20: CONSUMO FILA || Machine Learning Cubos
   RUNG wire#powerrail
      "CONSUMO_PRODUTO_LINHAS_EDI_ETR_DB"()
   END_RUNG
   RUNG wire#powerrail
      "DB_MachineLearnig_CUBOS_Instance"()
   END_RUNG
   // the same network as SCL:
   "CONSUMO_PRODUTO_LINHAS_EDI_ETR_DB"();   // "CONSUMO_PRODUTO_LINHAS_EDI_ETR"
   "DB_MachineLearnig_CUBOS_Instance"();   // "FB_MachineLearnig_CUBOS"
END_REGION

REGION Network 21: DIAGNOSTICO_PROFINET
   RUNG wire#powerrail
      "DIAGNOSTICO_PROFINET_DB"()
   END_RUNG
   // the same network as SCL:
   "DIAGNOSTICO_PROFINET_DB"();   // "DIAGNOSTICO_PROFINET"
END_REGION

REGION Network 22: Desvios
   RUNG wire#powerrail
      "FC15_DeviationManager"()
   END_RUNG
   // the same network as SCL:
   "FC15_DeviationManager"();
END_REGION

REGION Network 23: BSEND SEQUENCE NOW MD1
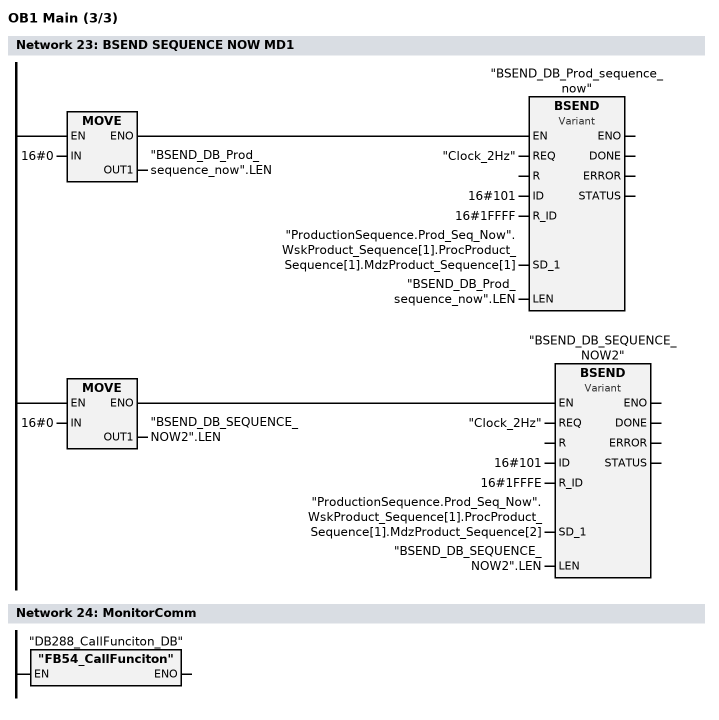
   RUNG wire#powerrail
      Move(in := 16#0, out1 => "BSEND_DB_Prod_sequence_now".LEN)
      { S7_Templates := "[ptr_type := Variant, id_type := CONN_PRG, r_id_type := CONN_R_ID]" } "BSEND_DB_Prod_sequence_now".BSEND(REQ := "Clock_2Hz", R :=, ID := 16#101, R_ID := 16#1FFFF, SD_1 := "ProductionSequence.Prod_Seq_Now".WskProduct_Sequence[1].ProcProduct_Sequence[1].MdzProduct_Sequence[1], LEN := "BSEND_DB_Prod_sequence_now".LEN, DONE =>, ERROR =>, STATUS =>)
   END_RUNG
   RUNG wire#powerrail
      Move(in := 16#0, out1 => "BSEND_DB_SEQUENCE_NOW2".LEN)
      { S7_Templates := "[ptr_type := Variant, id_type := CONN_PRG, r_id_type := CONN_R_ID]" } "BSEND_DB_SEQUENCE_NOW2".BSEND(REQ := "Clock_2Hz", R :=, ID := 16#101, R_ID := 16#1FFFE, SD_1 := "ProductionSequence.Prod_Seq_Now".WskProduct_Sequence[1].ProcProduct_Sequence[1].MdzProduct_Sequence[2], LEN := "BSEND_DB_SEQUENCE_NOW2".LEN, DONE =>, ERROR =>, STATUS =>)
   END_RUNG
   // the same network as SCL:
   "BSEND_DB_Prod_sequence_now".LEN := 16#0;
   "BSEND_DB_Prod_sequence_now"(REQ := "Clock_2Hz",   // BSEND
                           ID := 16#101,
                           R_ID := 16#1FFFF,
                           SD_1 := "ProductionSequence.Prod_Seq_Now".WskProduct_Sequence[1].ProcProduct_Sequence[1].MdzProduct_Sequence[1],
                           LEN := "BSEND_DB_Prod_sequence_now".LEN);
   "BSEND_DB_SEQUENCE_NOW2".LEN := 16#0;
   "BSEND_DB_SEQUENCE_NOW2"(REQ := "Clock_2Hz",   // BSEND
                           ID := 16#101,
                           R_ID := 16#1FFFE,
                           SD_1 := "ProductionSequence.Prod_Seq_Now".WskProduct_Sequence[1].ProcProduct_Sequence[1].MdzProduct_Sequence[2],
                           LEN := "BSEND_DB_SEQUENCE_NOW2".LEN);
END_REGION

REGION Network 24: MonitorComm
   RUNG wire#powerrail
      "DB288_CallFunciton_DB"()
   END_RUNG
   // the same network as SCL:
   "DB288_CallFunciton_DB"();   // "FB54_CallFunciton"
END_REGION
END_ORGANIZATION_BLOCK

FUNCTION "BYPASS DOS EQUIPAMENTOS" : Void   // FC12, LAD
{ S7_Optimized_Access := 'TRUE' }
// stored: SetENOAutomatically false
BEGIN

REGION Network 1: BYPASS GERAL E ESVAZIAMENTO DOS TRANSPORTADORES
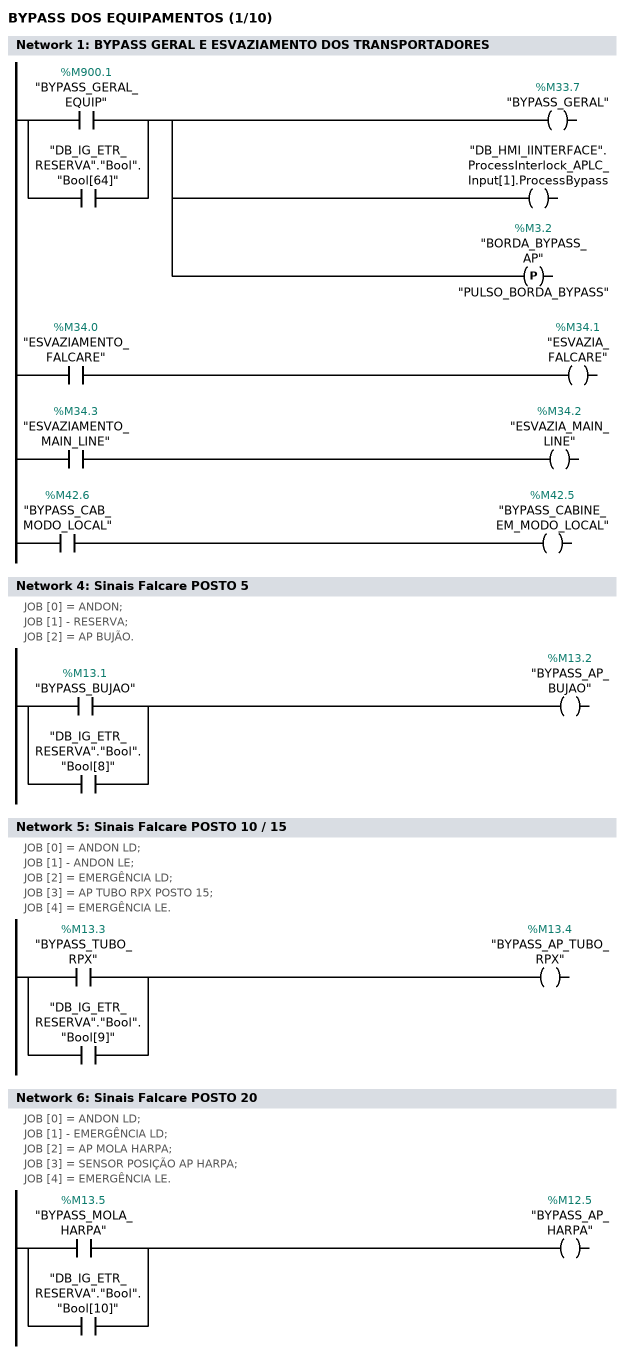
   "BYPASS_GERAL" := "BYPASS_GERAL_EQUIP" OR "DB_IG_ETR_RESERVA"."Bool"."Bool[64]";
   "DB_HMI_IINTERFACE".ProcessInterlock_APLC_Input[1].ProcessBypass := "BYPASS_GERAL";
   "BORDA_BYPASS_AP" := "BYPASS_GERAL" AND NOT "PULSO_BORDA_BYPASS";   // rising edge
   "PULSO_BORDA_BYPASS" := "BYPASS_GERAL";
   "ESVAZIA_FALCARE" := "ESVAZIAMENTO_FALCARE";
   "ESVAZIA_MAIN_LINE" := "ESVAZIAMENTO_MAIN_LINE";
   "BYPASS_CABINE_EM_MODO_LOCAL" := "BYPASS_CAB_MODO_LOCAL";
END_REGION

REGION Network 2: Sinais Falcare POSTO 1
   // JOB [0] = ANDON;
   // JOB [1] - EMERGÊNCIA;
END_REGION

REGION Network 3: Sinais Falcare VIVERK
   // JOB [0] = ANDON;
   // JOB [1] - EMERGÊNCIA;
END_REGION

REGION Network 4: Sinais Falcare POSTO 5
   // JOB [0] = ANDON;
   // JOB [1] - RESERVA;
   // JOB [2] = AP BUJÃO.
   RUNG wire#powerrail
      Contact( "BYPASS_BUJAO" )
      wire#w1
      Coil( "BYPASS_AP_BUJAO" )
   END_RUNG
   RUNG wire#powerrail
      Contact( "DB_IG_ETR_RESERVA"."Bool"."Bool[8]" )
   END_RUNG wire#w1
   // the same network as SCL:
   "BYPASS_AP_BUJAO" := "BYPASS_BUJAO" OR "DB_IG_ETR_RESERVA"."Bool"."Bool[8]";
END_REGION

REGION Network 5: Sinais Falcare POSTO 10 / 15
   // JOB [0] = ANDON LD;
   // JOB [1] - ANDON LE;
   // JOB [2] = EMERGÊNCIA LD;
   // JOB [3] = AP TUBO RPX POSTO 15;
   // JOB [4] = EMERGÊNCIA LE.
   RUNG wire#powerrail
      Contact( "BYPASS_TUBO_RPX" )
      wire#w1
      Coil( "BYPASS_AP_TUBO_RPX" )
   END_RUNG
   RUNG wire#powerrail
      Contact( "DB_IG_ETR_RESERVA"."Bool"."Bool[9]" )
   END_RUNG wire#w1
   // the same network as SCL:
   "BYPASS_AP_TUBO_RPX" := "BYPASS_TUBO_RPX" OR "DB_IG_ETR_RESERVA"."Bool"."Bool[9]";
END_REGION

REGION Network 6: Sinais Falcare POSTO 20
   // JOB [0] = ANDON LD;
   // JOB [1] - EMERGÊNCIA LD;
   // JOB [2] = AP MOLA HARPA;
   // JOB [3] = SENSOR POSIÇÃO AP HARPA;
   // JOB [4] = EMERGÊNCIA LE.
   RUNG wire#powerrail
      Contact( "BYPASS_MOLA_HARPA" )
      wire#w1
      Coil( "BYPASS_AP_HARPA" )
   END_RUNG
   RUNG wire#powerrail
      Contact( "DB_IG_ETR_RESERVA"."Bool"."Bool[10]" )
   END_RUNG wire#w1
   // the same network as SCL:
   "BYPASS_AP_HARPA" := "BYPASS_MOLA_HARPA" OR "DB_IG_ETR_RESERVA"."Bool"."Bool[10]";
END_REGION

REGION Network 7: Sinais Falcare POSTO 30
   // JOB [0] = ANDON LD;
   // JOB [1] = ANDON LE;
   // JOB [2] = EMERGENCIA;
   // JOB [3] = AP DA CARCAÇA;
   // JOB [4] = POSIÇÃO TALHA DIF.
   // JOB [5] = PY JUNTA.
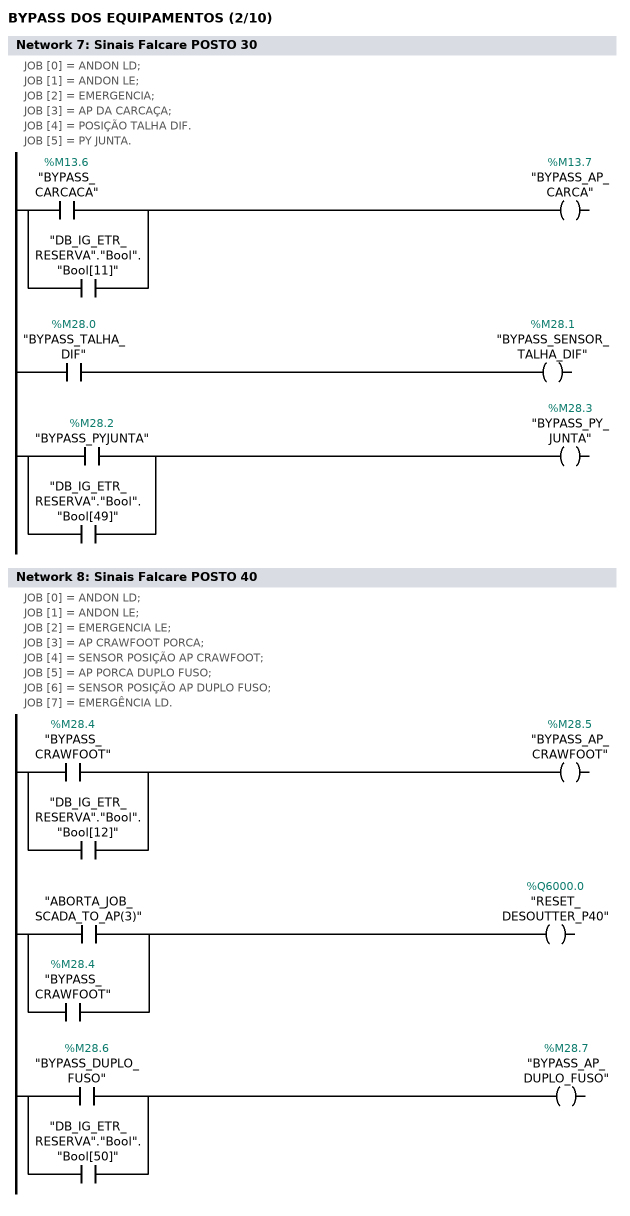
   RUNG wire#powerrail
      Contact( "BYPASS_CARCACA" )
      wire#w1
      Coil( "BYPASS_AP_CARCA" )
   END_RUNG
   RUNG wire#powerrail
      Contact( "DB_IG_ETR_RESERVA"."Bool"."Bool[11]" )
   END_RUNG wire#w1
   RUNG wire#powerrail
      Contact( "BYPASS_TALHA_DIF" )
      Coil( "BYPASS_SENSOR_TALHA_DIF" )
   END_RUNG
   RUNG wire#powerrail
      Contact( "BYPASS_PYJUNTA" )
      wire#w2
      Coil( "BYPASS_PY_JUNTA" )
   END_RUNG
   RUNG wire#powerrail
      Contact( "DB_IG_ETR_RESERVA"."Bool"."Bool[49]" )
   END_RUNG wire#w2
   // the same network as SCL:
   "BYPASS_AP_CARCA" := "BYPASS_CARCACA" OR "DB_IG_ETR_RESERVA"."Bool"."Bool[11]";
   "BYPASS_SENSOR_TALHA_DIF" := "BYPASS_TALHA_DIF";
   "BYPASS_PY_JUNTA" := "BYPASS_PYJUNTA" OR "DB_IG_ETR_RESERVA"."Bool"."Bool[49]";
END_REGION

REGION Network 8: Sinais Falcare POSTO 40
   // JOB [0] = ANDON LD;
   // JOB [1] = ANDON LE;
   // JOB [2] = EMERGENCIA LE;
   // JOB [3] = AP CRAWFOOT PORCA;
   // JOB [4] = SENSOR POSIÇÃO AP CRAWFOOT;
   // JOB [5] = AP PORCA DUPLO FUSO;
   // JOB [6] = SENSOR POSIÇÃO AP DUPLO FUSO;
   // JOB [7] = EMERGÊNCIA LD.
   RUNG wire#powerrail
      Contact( "BYPASS_CRAWFOOT" )
      wire#w1
      Coil( "BYPASS_AP_CRAWFOOT" )
   END_RUNG
   RUNG wire#powerrail
      Contact( "DB_IG_ETR_RESERVA"."Bool"."Bool[12]" )
   END_RUNG wire#w1
   RUNG wire#powerrail
      Contact( "ABORTA_JOB_SCADA_TO_AP(3)" )
      wire#w2
      Coil( "RESET_DESOUTTER_P40" )
   END_RUNG
   RUNG wire#powerrail
      Contact( "BYPASS_CRAWFOOT" )
   END_RUNG wire#w2
   RUNG wire#powerrail
      Contact( "BYPASS_DUPLO_FUSO" )
      wire#w3
      Coil( "BYPASS_AP_DUPLO_FUSO" )
   END_RUNG
   RUNG wire#powerrail
      Contact( "DB_IG_ETR_RESERVA"."Bool"."Bool[50]" )
   END_RUNG wire#w3
   // the same network as SCL:
   "BYPASS_AP_CRAWFOOT" := "BYPASS_CRAWFOOT" OR "DB_IG_ETR_RESERVA"."Bool"."Bool[12]";
   "RESET_DESOUTTER_P40" := "ABORTA_JOB_SCADA_TO_AP(3)" OR "BYPASS_CRAWFOOT";
   "BYPASS_AP_DUPLO_FUSO" := "BYPASS_DUPLO_FUSO" OR "DB_IG_ETR_RESERVA"."Bool"."Bool[50]";
END_REGION

REGION Network 9: Sinais Falcare POSTO 50 /55
   // JOB [0] = ANDON;
   // JOB [1] = EMERGENCIA;
   // JOB [2] = AP PORCA ESCONDIDA;
   // JOB [3] = SENSOR POSIÇÃO AP PORCA ESCONDIDA;
   // JOB [4] = AP PORCA SUPORTE DO CILINDRO;
   // JOB [5] = SENSOR POSIÇÃO AP SUPORTE DO CILINDRO;
   // JOB [6] = ANDON LD.
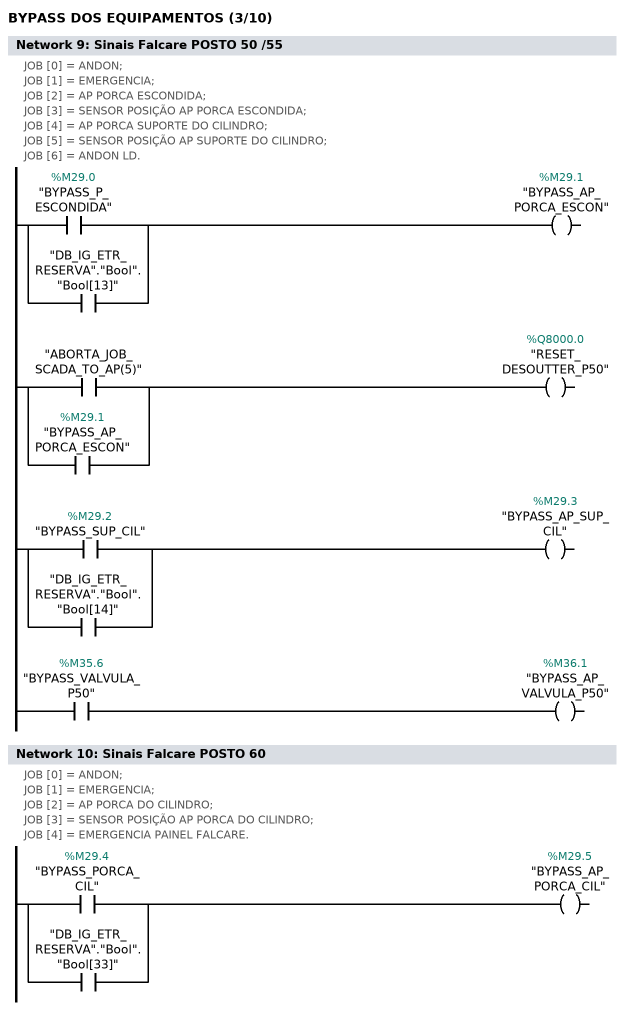
   RUNG wire#powerrail
      Contact( "BYPASS_P_ESCONDIDA" )
      wire#w1
      Coil( "BYPASS_AP_PORCA_ESCON" )
   END_RUNG
   RUNG wire#powerrail
      Contact( "DB_IG_ETR_RESERVA"."Bool"."Bool[13]" )
   END_RUNG wire#w1
   RUNG wire#powerrail
      Contact( "ABORTA_JOB_SCADA_TO_AP(5)" )
      wire#w2
      Coil( "RESET_DESOUTTER_P50" )
   END_RUNG
   RUNG wire#powerrail
      Contact( "BYPASS_AP_PORCA_ESCON" )
   END_RUNG wire#w2
   RUNG wire#powerrail
      Contact( "BYPASS_SUP_CIL" )
      wire#w3
      Coil( "BYPASS_AP_SUP_CIL" )
   END_RUNG
   RUNG wire#powerrail
      Contact( "DB_IG_ETR_RESERVA"."Bool"."Bool[14]" )
   END_RUNG wire#w3
   RUNG wire#powerrail
      Contact( "BYPASS_VALVULA_P50" )
      Coil( "BYPASS_AP_VALVULA_P50" )
   END_RUNG
   // the same network as SCL:
   "BYPASS_AP_PORCA_ESCON" := "BYPASS_P_ESCONDIDA" OR "DB_IG_ETR_RESERVA"."Bool"."Bool[13]";
   "RESET_DESOUTTER_P50" := "ABORTA_JOB_SCADA_TO_AP(5)" OR "BYPASS_AP_PORCA_ESCON";
   "BYPASS_AP_SUP_CIL" := "BYPASS_SUP_CIL" OR "DB_IG_ETR_RESERVA"."Bool"."Bool[14]";
   "BYPASS_AP_VALVULA_P50" := "BYPASS_VALVULA_P50";
END_REGION

REGION Network 10: Sinais Falcare POSTO 60
   // JOB [0] = ANDON;
   // JOB [1] = EMERGENCIA;
   // JOB [2] = AP PORCA DO CILINDRO;
   // JOB [3] = SENSOR POSIÇÃO AP PORCA DO CILINDRO;
   // JOB [4] = EMERGENCIA PAINEL FALCARE.
   RUNG wire#powerrail
      Contact( "BYPASS_PORCA_CIL" )
      wire#w1
      Coil( "BYPASS_AP_PORCA_CIL" )
   END_RUNG
   RUNG wire#powerrail
      Contact( "DB_IG_ETR_RESERVA"."Bool"."Bool[33]" )
   END_RUNG wire#w1
   // the same network as SCL:
   "BYPASS_AP_PORCA_CIL" := "BYPASS_PORCA_CIL" OR "DB_IG_ETR_RESERVA"."Bool"."Bool[33]";
END_REGION

REGION Network 11: Sinais Main Line POSTO 70 / 75
   // \\ JOB [0] - ANDON
END_REGION

REGION Network 12: Sinais Main Line POSTO 80
   // JOB [0]=- ANDON;
   // JOB [1] = EMERGÊNCIA;
   // JOB [2] = AP SUP FREIO;
   // JOB [3] = PY EIXO EXCENTRICO;
   // JOB [4] = PY CUBO DISCO
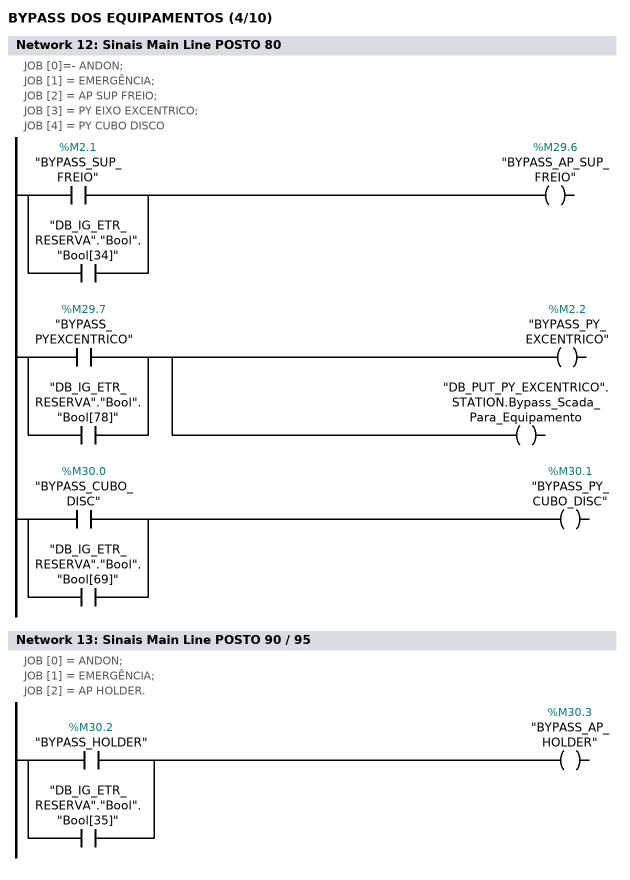
   RUNG wire#powerrail
      Contact( "BYPASS_SUP_FREIO" )
      wire#w1
      Coil( "BYPASS_AP_SUP_FREIO" )
   END_RUNG
   RUNG wire#powerrail
      Contact( "DB_IG_ETR_RESERVA"."Bool"."Bool[34]" )
   END_RUNG wire#w1
   RUNG wire#powerrail
      Contact( "BYPASS_PYEXCENTRICO" )
      wire#w2
      Coil( "BYPASS_PY_EXCENTRICO" )
   END_RUNG
   RUNG wire#powerrail
      Contact( "DB_IG_ETR_RESERVA"."Bool"."Bool[78]" )
   END_RUNG wire#w2
   RUNG wire#w2
      Coil( "DB_PUT_PY_EXCENTRICO".STATION.Bypass_Scada_Para_Equipamento )
   END_RUNG
   RUNG wire#powerrail
      Contact( "BYPASS_CUBO_DISC" )
      wire#w3
      Coil( "BYPASS_PY_CUBO_DISC" )
   END_RUNG
   RUNG wire#powerrail
      Contact( "DB_IG_ETR_RESERVA"."Bool"."Bool[69]" )
   END_RUNG wire#w3
   // the same network as SCL:
   "BYPASS_AP_SUP_FREIO" := "BYPASS_SUP_FREIO" OR "DB_IG_ETR_RESERVA"."Bool"."Bool[34]";
   "BYPASS_PY_EXCENTRICO" := "BYPASS_PYEXCENTRICO" OR "DB_IG_ETR_RESERVA"."Bool"."Bool[78]";
   "DB_PUT_PY_EXCENTRICO".STATION.Bypass_Scada_Para_Equipamento := "BYPASS_PY_EXCENTRICO";
   "BYPASS_PY_CUBO_DISC" := "BYPASS_CUBO_DISC" OR "DB_IG_ETR_RESERVA"."Bool"."Bool[69]";
END_REGION

REGION Network 13: Sinais Main Line POSTO 90 / 95
   // JOB [0] = ANDON;
   // JOB [1] = EMERGÊNCIA;
   // JOB [2] = AP HOLDER.
   RUNG wire#powerrail
      Contact( "BYPASS_HOLDER" )
      wire#w1
      Coil( "BYPASS_AP_HOLDER" )
   END_RUNG
   RUNG wire#powerrail
      Contact( "DB_IG_ETR_RESERVA"."Bool"."Bool[35]" )
   END_RUNG wire#w1
   // the same network as SCL:
   "BYPASS_AP_HOLDER" := "BYPASS_HOLDER" OR "DB_IG_ETR_RESERVA"."Bool"."Bool[35]";
END_REGION

REGION Network 14: Sinais Main Line POSTO100 /105
   // JOB [0] = ANDON;
   // JOB [1] = EMERGÊNCIA;
   // JOB [2] = AP CALIPER;
   // JOB [3] = PY CUBO TAMBOR;
   // JOB [4] = ANDON P105;
   // JOB [5] = AP HASTE ALAVANCA
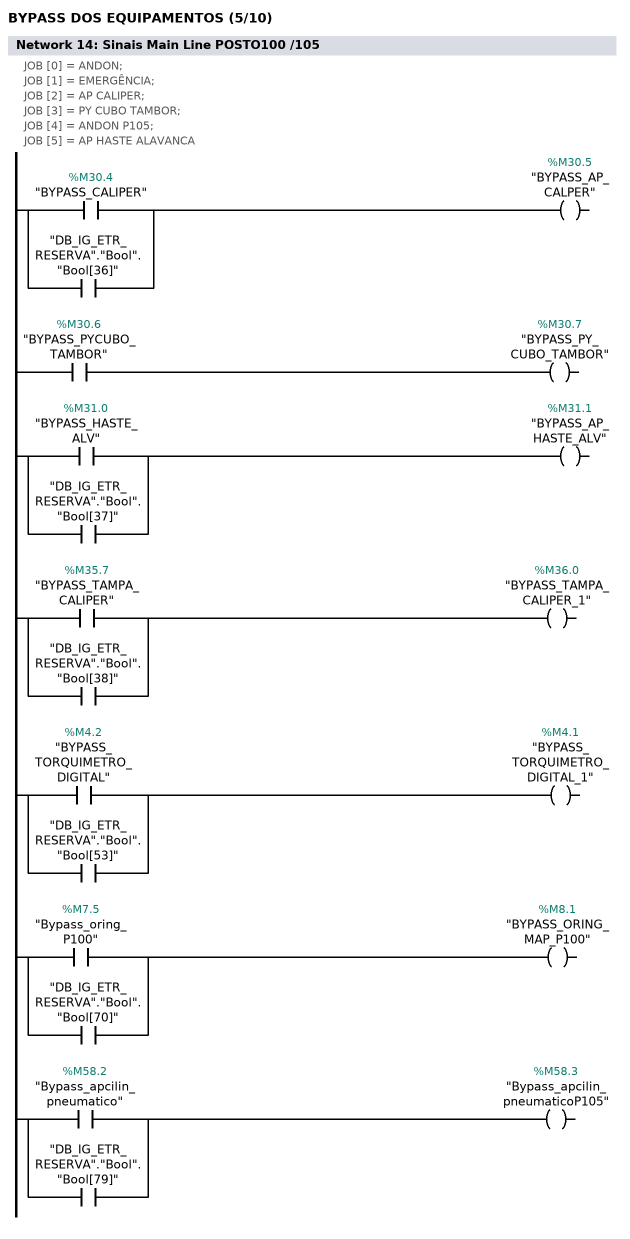
   RUNG wire#powerrail
      Contact( "BYPASS_CALIPER" )
      wire#w1
      Coil( "BYPASS_AP_CALPER" )
   END_RUNG
   RUNG wire#powerrail
      Contact( "DB_IG_ETR_RESERVA"."Bool"."Bool[36]" )
   END_RUNG wire#w1
   RUNG wire#powerrail
      Contact( "BYPASS_PYCUBO_TAMBOR" )
      Coil( "BYPASS_PY_CUBO_TAMBOR" )
   END_RUNG
   RUNG wire#powerrail
      Contact( "BYPASS_HASTE_ALV" )
      wire#w2
      Coil( "BYPASS_AP_HASTE_ALV" )
   END_RUNG
   RUNG wire#powerrail
      Contact( "DB_IG_ETR_RESERVA"."Bool"."Bool[37]" )
   END_RUNG wire#w2
   RUNG wire#powerrail
      Contact( "BYPASS_TAMPA_CALIPER" )
      wire#w3
      Coil( "BYPASS_TAMPA_CALIPER_1" )
   END_RUNG
   RUNG wire#powerrail
      Contact( "DB_IG_ETR_RESERVA"."Bool"."Bool[38]" )
   END_RUNG wire#w3
   RUNG wire#powerrail
      Contact( "BYPASS_TORQUIMETRO_DIGITAL" )
      wire#w4
      Coil( "BYPASS_TORQUIMETRO_DIGITAL_1" )
   END_RUNG
   RUNG wire#powerrail
      Contact( "DB_IG_ETR_RESERVA"."Bool"."Bool[53]" )
   END_RUNG wire#w4
   RUNG wire#powerrail
      Contact( "Bypass_oring_P100" )
      wire#w5
      Coil( "BYPASS_ORING_MAP_P100" )
   END_RUNG
   RUNG wire#powerrail
      Contact( "DB_IG_ETR_RESERVA"."Bool"."Bool[70]" )
   END_RUNG wire#w5
   RUNG wire#powerrail
      Contact( "Bypass_apcilin_pneumatico" )
      wire#w6
      Coil( "Bypass_apcilin_pneumaticoP105" )
   END_RUNG
   RUNG wire#powerrail
      Contact( "DB_IG_ETR_RESERVA"."Bool"."Bool[79]" )
   END_RUNG wire#w6
   // the same network as SCL:
   "BYPASS_AP_CALPER" := "BYPASS_CALIPER" OR "DB_IG_ETR_RESERVA"."Bool"."Bool[36]";
   "BYPASS_PY_CUBO_TAMBOR" := "BYPASS_PYCUBO_TAMBOR";
   "BYPASS_AP_HASTE_ALV" := "BYPASS_HASTE_ALV" OR "DB_IG_ETR_RESERVA"."Bool"."Bool[37]";
   "BYPASS_TAMPA_CALIPER_1" := "BYPASS_TAMPA_CALIPER" OR "DB_IG_ETR_RESERVA"."Bool"."Bool[38]";
   "BYPASS_TORQUIMETRO_DIGITAL_1" := "BYPASS_TORQUIMETRO_DIGITAL" OR "DB_IG_ETR_RESERVA"."Bool"."Bool[53]";
   "BYPASS_ORING_MAP_P100" := "Bypass_oring_P100" OR "DB_IG_ETR_RESERVA"."Bool"."Bool[70]";
   "Bypass_apcilin_pneumaticoP105" := "Bypass_apcilin_pneumatico" OR "DB_IG_ETR_RESERVA"."Bool"."Bool[79]";
END_REGION

REGION Network 15: Sinais Main Line POSTO110 /115
   // JOB [0] = ANDON;
   // JOB [1] = SEG. BLOQUEIO CLP;
   // JOB [2] = AP CUBO;
   // JOB [3] = ANDON P115;
   // JOB [4] = CRAVADOR.
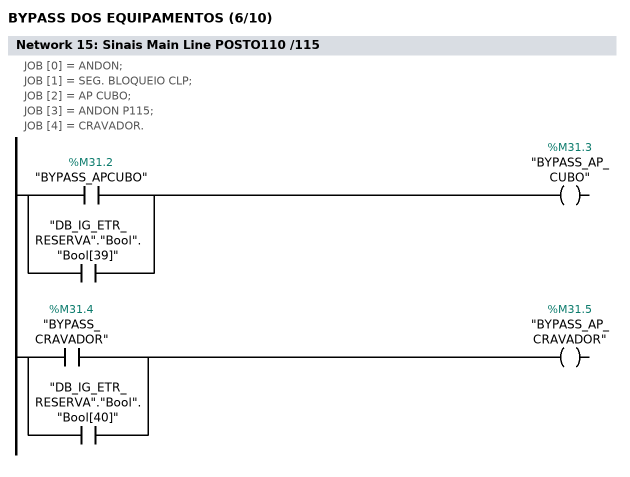
   RUNG wire#powerrail
      Contact( "BYPASS_APCUBO" )
      wire#w1
      Coil( "BYPASS_AP_CUBO" )
   END_RUNG
   RUNG wire#powerrail
      Contact( "DB_IG_ETR_RESERVA"."Bool"."Bool[39]" )
   END_RUNG wire#w1
   RUNG wire#powerrail
      Contact( "BYPASS_CRAVADOR" )
      wire#w2
      Coil( "BYPASS_AP_CRAVADOR" )
   END_RUNG
   RUNG wire#powerrail
      Contact( "DB_IG_ETR_RESERVA"."Bool"."Bool[40]" )
   END_RUNG wire#w2
   // the same network as SCL:
   "BYPASS_AP_CUBO" := "BYPASS_APCUBO" OR "DB_IG_ETR_RESERVA"."Bool"."Bool[39]";
   "BYPASS_AP_CRAVADOR" := "BYPASS_CRAVADOR" OR "DB_IG_ETR_RESERVA"."Bool"."Bool[40]";
END_REGION

REGION Network 16: Sinais Main Line POSTO120 /125
   // JOB [0] = ANDON;
   // JOB [1] - EMERGÊNCIA;
   // JOB [2] = AP INDICADOR;
   // JOB [3] = AP VALVULA;
   // JOB [4] = PY HELGE;
   // JOB [5] - ANDON P125;
   // JOB [6] - AP PORCA TERMINAL;
   // JOB [7] - AP FILTRO OLEO.
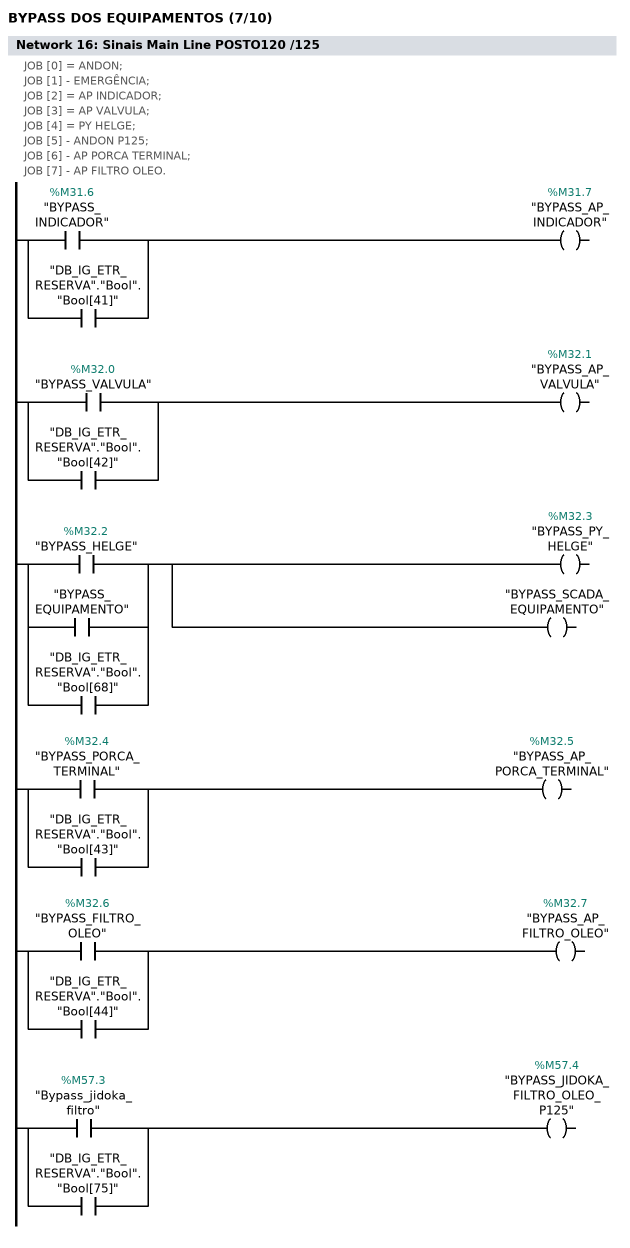
   RUNG wire#powerrail
      Contact( "BYPASS_INDICADOR" )
      wire#w1
      Coil( "BYPASS_AP_INDICADOR" )
   END_RUNG
   RUNG wire#powerrail
      Contact( "DB_IG_ETR_RESERVA"."Bool"."Bool[41]" )
   END_RUNG wire#w1
   RUNG wire#powerrail
      Contact( "BYPASS_VALVULA" )
      wire#w2
      Coil( "BYPASS_AP_VALVULA" )
   END_RUNG
   RUNG wire#powerrail
      Contact( "DB_IG_ETR_RESERVA"."Bool"."Bool[42]" )
   END_RUNG wire#w2
   RUNG wire#powerrail
      Contact( "BYPASS_HELGE" )
      wire#w3
      Coil( "BYPASS_PY_HELGE" )
   END_RUNG
   RUNG wire#powerrail
      Contact( "BYPASS_EQUIPAMENTO" )
   END_RUNG wire#w3
   RUNG wire#powerrail
      Contact( "DB_IG_ETR_RESERVA"."Bool"."Bool[68]" )
   END_RUNG wire#w3
   RUNG wire#w3
      Coil( "BYPASS_SCADA_EQUIPAMENTO" )
   END_RUNG
   RUNG wire#powerrail
      Contact( "BYPASS_PORCA_TERMINAL" )
      wire#w4
      Coil( "BYPASS_AP_PORCA_TERMINAL" )
   END_RUNG
   RUNG wire#powerrail
      Contact( "DB_IG_ETR_RESERVA"."Bool"."Bool[43]" )
   END_RUNG wire#w4
   RUNG wire#powerrail
      Contact( "BYPASS_FILTRO_OLEO" )
      wire#w5
      Coil( "BYPASS_AP_FILTRO_OLEO" )
   END_RUNG
   RUNG wire#powerrail
      Contact( "DB_IG_ETR_RESERVA"."Bool"."Bool[44]" )
   END_RUNG wire#w5
   RUNG wire#powerrail
      Contact( "Bypass_jidoka_filtro" )
      wire#w6
      Coil( "BYPASS_JIDOKA_FILTRO_OLEO_P125" )
   END_RUNG
   RUNG wire#powerrail
      Contact( "DB_IG_ETR_RESERVA"."Bool"."Bool[75]" )
   END_RUNG wire#w6
   // the same network as SCL:
   "BYPASS_AP_INDICADOR" := "BYPASS_INDICADOR" OR "DB_IG_ETR_RESERVA"."Bool"."Bool[41]";
   "BYPASS_AP_VALVULA" := "BYPASS_VALVULA" OR "DB_IG_ETR_RESERVA"."Bool"."Bool[42]";
   "BYPASS_PY_HELGE" := "BYPASS_HELGE" OR "BYPASS_EQUIPAMENTO" OR "DB_IG_ETR_RESERVA"."Bool"."Bool[68]";
   "BYPASS_SCADA_EQUIPAMENTO" := "BYPASS_PY_HELGE";
   "BYPASS_AP_PORCA_TERMINAL" := "BYPASS_PORCA_TERMINAL" OR "DB_IG_ETR_RESERVA"."Bool"."Bool[43]";
   "BYPASS_AP_FILTRO_OLEO" := "BYPASS_FILTRO_OLEO" OR "DB_IG_ETR_RESERVA"."Bool"."Bool[44]";
   "BYPASS_JIDOKA_FILTRO_OLEO_P125" := "Bypass_jidoka_filtro" OR "DB_IG_ETR_RESERVA"."Bool"."Bool[75]";
END_REGION

REGION Network 17: Sinais Main Line POSTO130
   // JOB [0] = ANDON;
   // JOB [1] = AP REDUÇÃO;
   // JOB [2] - AP FALNGE
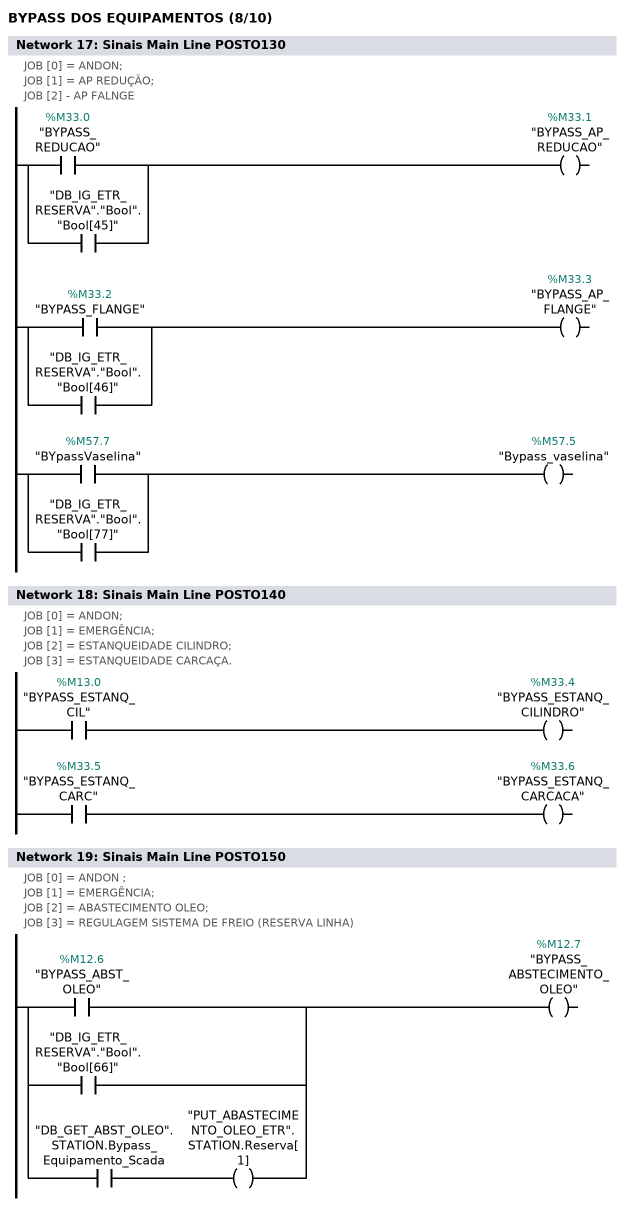
   RUNG wire#powerrail
      Contact( "BYPASS_REDUCAO" )
      wire#w1
      Coil( "BYPASS_AP_REDUCAO" )
   END_RUNG
   RUNG wire#powerrail
      Contact( "DB_IG_ETR_RESERVA"."Bool"."Bool[45]" )
   END_RUNG wire#w1
   RUNG wire#powerrail
      Contact( "BYPASS_FLANGE" )
      wire#w2
      Coil( "BYPASS_AP_FLANGE" )
   END_RUNG
   RUNG wire#powerrail
      Contact( "DB_IG_ETR_RESERVA"."Bool"."Bool[46]" )
   END_RUNG wire#w2
   RUNG wire#powerrail
      Contact( "BYpassVaselina" )
      wire#w3
      Coil( "Bypass_vaselina" )
   END_RUNG
   RUNG wire#powerrail
      Contact( "DB_IG_ETR_RESERVA"."Bool"."Bool[77]" )
   END_RUNG wire#w3
   // the same network as SCL:
   "BYPASS_AP_REDUCAO" := "BYPASS_REDUCAO" OR "DB_IG_ETR_RESERVA"."Bool"."Bool[45]";
   "BYPASS_AP_FLANGE" := "BYPASS_FLANGE" OR "DB_IG_ETR_RESERVA"."Bool"."Bool[46]";
   "Bypass_vaselina" := "BYpassVaselina" OR "DB_IG_ETR_RESERVA"."Bool"."Bool[77]";
END_REGION

REGION Network 18: Sinais Main Line POSTO140
   // JOB [0] = ANDON;
   // JOB [1] = EMERGÊNCIA;
   // JOB [2] = ESTANQUEIDADE CILINDRO;
   // JOB [3] = ESTANQUEIDADE CARCAÇA.
   RUNG wire#powerrail
      Contact( "BYPASS_ESTANQ_CIL" )
      Coil( "BYPASS_ESTANQ_CILINDRO" )
   END_RUNG
   RUNG wire#powerrail
      Contact( "BYPASS_ESTANQ_CARC" )
      Coil( "BYPASS_ESTANQ_CARCACA" )
   END_RUNG
   // the same network as SCL:
   "BYPASS_ESTANQ_CILINDRO" := "BYPASS_ESTANQ_CIL";
   "BYPASS_ESTANQ_CARCACA" := "BYPASS_ESTANQ_CARC";
END_REGION

REGION Network 19: Sinais Main Line POSTO150
   // JOB [0] = ANDON ;
   // JOB [1] = EMERGÊNCIA;
   // JOB [2] = ABASTECIMENTO OLEO;
   // JOB [3] = REGULAGEM SISTEMA DE FREIO (RESERVA LINHA)
   RUNG wire#powerrail
      Contact( "BYPASS_ABST_OLEO" )
      wire#w1
      Coil( "BYPASS_ABSTECIMENTO_OLEO" )
   END_RUNG
   RUNG wire#powerrail
      Contact( "DB_IG_ETR_RESERVA"."Bool"."Bool[66]" )
   END_RUNG wire#w1
   RUNG wire#powerrail
      Contact( "DB_GET_ABST_OLEO".STATION.Bypass_Equipamento_Scada )
      Coil( "PUT_ABASTECIMENTO_OLEO_ETR".STATION.Reserva[1] )
   END_RUNG wire#w1
   // the same network as SCL:
   "PUT_ABASTECIMENTO_OLEO_ETR".STATION.Reserva[1] := "DB_GET_ABST_OLEO".STATION.Bypass_Equipamento_Scada;
   "BYPASS_ABSTECIMENTO_OLEO" := "BYPASS_ABST_OLEO" OR "DB_IG_ETR_RESERVA"."Bool"."Bool[66]" OR "DB_GET_ABST_OLEO".STATION.Bypass_Equipamento_Scada;
END_REGION

REGION Network 20: Sinais Main Line Q.G
   // JOB [0] = ANDON;
   // JOB [1] = EMERGÊNCIA;
   // JOB [2] - EIXO PENDURADO;
   // JOB [3] - GAP PRESENTE CAB;
   // JOB [4] - GAP PRESENTE TAKT
END_REGION

REGION Network 21: Sinais Main Line EXPEDIÇÃO
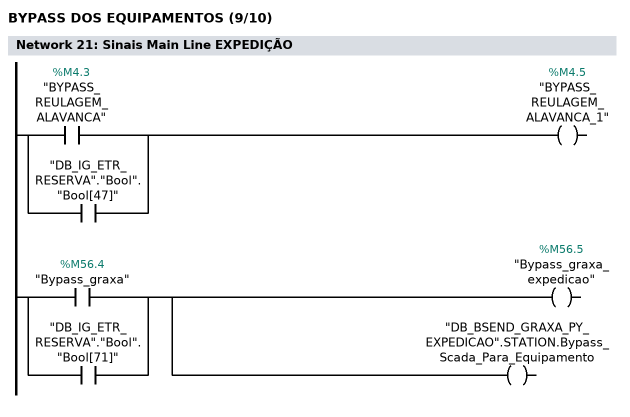
   RUNG wire#powerrail
      Contact( "BYPASS_REULAGEM_ALAVANCA" )
      wire#w1
      Coil( "BYPASS_REULAGEM_ALAVANCA_1" )
   END_RUNG
   RUNG wire#powerrail
      Contact( "DB_IG_ETR_RESERVA"."Bool"."Bool[47]" )
   END_RUNG wire#w1
   RUNG wire#powerrail
      Contact( "Bypass_graxa" )
      wire#w2
      Coil( "Bypass_graxa_expedicao" )
   END_RUNG
   RUNG wire#powerrail
      Contact( "DB_IG_ETR_RESERVA"."Bool"."Bool[71]" )
   END_RUNG wire#w2
   RUNG wire#w2
      Coil( "DB_BSEND_GRAXA_PY_EXPEDICAO".STATION.Bypass_Scada_Para_Equipamento )
   END_RUNG
   // the same network as SCL:
   "BYPASS_REULAGEM_ALAVANCA_1" := "BYPASS_REULAGEM_ALAVANCA" OR "DB_IG_ETR_RESERVA"."Bool"."Bool[47]";
   "Bypass_graxa_expedicao" := "Bypass_graxa" OR "DB_IG_ETR_RESERVA"."Bool"."Bool[71]";
   "DB_BSEND_GRAXA_PY_EXPEDICAO".STATION.Bypass_Scada_Para_Equipamento := "Bypass_graxa_expedicao";
END_REGION

REGION Network 22: BYPASS STATIONS
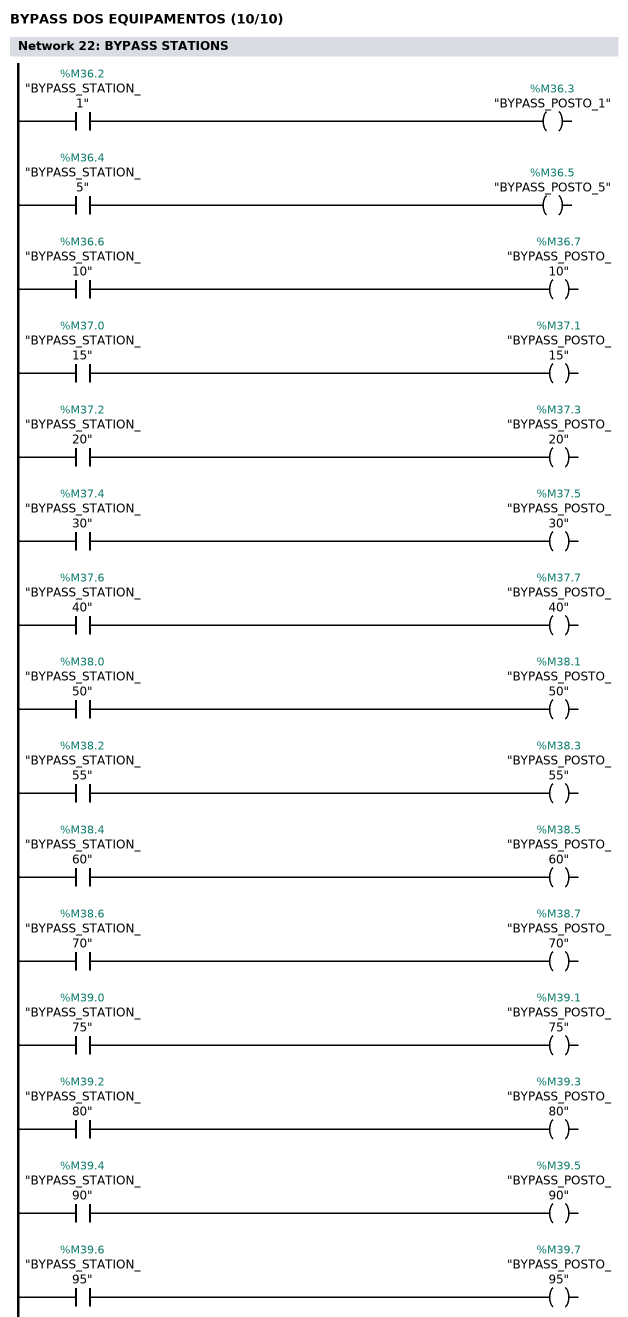
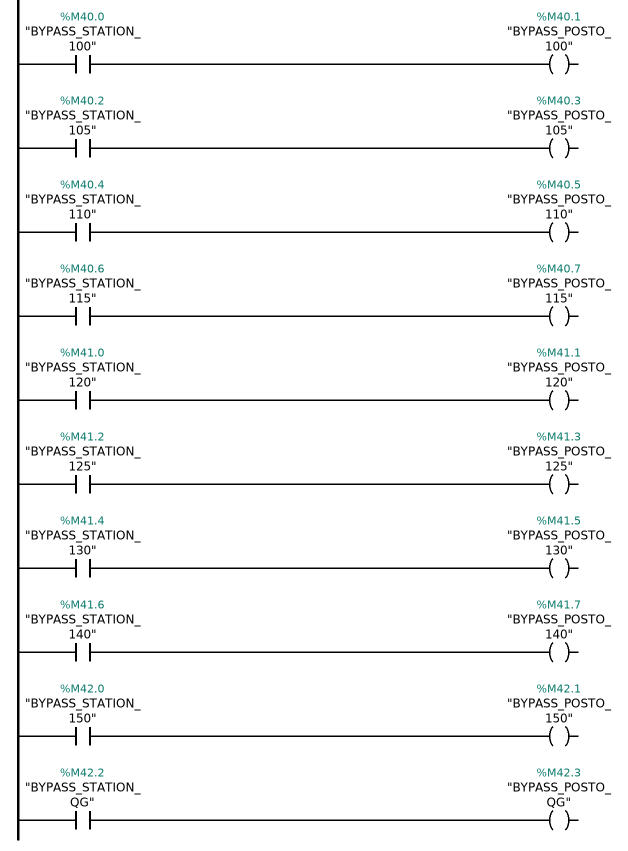
   RUNG wire#powerrail
      Contact( "BYPASS_STATION_1" )
      Coil( "BYPASS_POSTO_1" )
   END_RUNG
   RUNG wire#powerrail
      Contact( "BYPASS_STATION_5" )
      Coil( "BYPASS_POSTO_5" )
   END_RUNG
   RUNG wire#powerrail
      Contact( "BYPASS_STATION_10" )
      Coil( "BYPASS_POSTO_10" )
   END_RUNG
   RUNG wire#powerrail
      Contact( "BYPASS_STATION_15" )
      Coil( "BYPASS_POSTO_15" )
   END_RUNG
   RUNG wire#powerrail
      Contact( "BYPASS_STATION_20" )
      Coil( "BYPASS_POSTO_20" )
   END_RUNG
   RUNG wire#powerrail
      Contact( "BYPASS_STATION_30" )
      Coil( "BYPASS_POSTO_30" )
   END_RUNG
   RUNG wire#powerrail
      Contact( "BYPASS_STATION_40" )
      Coil( "BYPASS_POSTO_40" )
   END_RUNG
   RUNG wire#powerrail
      Contact( "BYPASS_STATION_50" )
      Coil( "BYPASS_POSTO_50" )
   END_RUNG
   RUNG wire#powerrail
      Contact( "BYPASS_STATION_55" )
      Coil( "BYPASS_POSTO_55" )
   END_RUNG
   RUNG wire#powerrail
      Contact( "BYPASS_STATION_60" )
      Coil( "BYPASS_POSTO_60" )
   END_RUNG
   RUNG wire#powerrail
      Contact( "BYPASS_STATION_70" )
      Coil( "BYPASS_POSTO_70" )
   END_RUNG
   RUNG wire#powerrail
      Contact( "BYPASS_STATION_75" )
      Coil( "BYPASS_POSTO_75" )
   END_RUNG
   RUNG wire#powerrail
      Contact( "BYPASS_STATION_80" )
      Coil( "BYPASS_POSTO_80" )
   END_RUNG
   RUNG wire#powerrail
      Contact( "BYPASS_STATION_90" )
      Coil( "BYPASS_POSTO_90" )
   END_RUNG
   RUNG wire#powerrail
      Contact( "BYPASS_STATION_95" )
      Coil( "BYPASS_POSTO_95" )
   END_RUNG
   RUNG wire#powerrail
      Contact( "BYPASS_STATION_100" )
      Coil( "BYPASS_POSTO_100" )
   END_RUNG
   RUNG wire#powerrail
      Contact( "BYPASS_STATION_105" )
      Coil( "BYPASS_POSTO_105" )
   END_RUNG
   RUNG wire#powerrail
      Contact( "BYPASS_STATION_110" )
      Coil( "BYPASS_POSTO_110" )
   END_RUNG
   RUNG wire#powerrail
      Contact( "BYPASS_STATION_115" )
      Coil( "BYPASS_POSTO_115" )
   END_RUNG
   RUNG wire#powerrail
      Contact( "BYPASS_STATION_120" )
      Coil( "BYPASS_POSTO_120" )
   END_RUNG
   RUNG wire#powerrail
      Contact( "BYPASS_STATION_125" )
      Coil( "BYPASS_POSTO_125" )
   END_RUNG
   RUNG wire#powerrail
      Contact( "BYPASS_STATION_130" )
      Coil( "BYPASS_POSTO_130" )
   END_RUNG
   RUNG wire#powerrail
      Contact( "BYPASS_STATION_140" )
      Coil( "BYPASS_POSTO_140" )
   END_RUNG
   RUNG wire#powerrail
      Contact( "BYPASS_STATION_150" )
      Coil( "BYPASS_POSTO_150" )
   END_RUNG
   RUNG wire#powerrail
      Contact( "BYPASS_STATION_QG" )
      Coil( "BYPASS_POSTO_QG" )
   END_RUNG
   // the same network as SCL:
   "BYPASS_POSTO_1" := "BYPASS_STATION_1";
   "BYPASS_POSTO_5" := "BYPASS_STATION_5";
   "BYPASS_POSTO_10" := "BYPASS_STATION_10";
   "BYPASS_POSTO_15" := "BYPASS_STATION_15";
   "BYPASS_POSTO_20" := "BYPASS_STATION_20";
   "BYPASS_POSTO_30" := "BYPASS_STATION_30";
   "BYPASS_POSTO_40" := "BYPASS_STATION_40";
   "BYPASS_POSTO_50" := "BYPASS_STATION_50";
   "BYPASS_POSTO_55" := "BYPASS_STATION_55";
   "BYPASS_POSTO_60" := "BYPASS_STATION_60";
   "BYPASS_POSTO_70" := "BYPASS_STATION_70";
   "BYPASS_POSTO_75" := "BYPASS_STATION_75";
   "BYPASS_POSTO_80" := "BYPASS_STATION_80";
   "BYPASS_POSTO_90" := "BYPASS_STATION_90";
   "BYPASS_POSTO_95" := "BYPASS_STATION_95";
   "BYPASS_POSTO_100" := "BYPASS_STATION_100";
   "BYPASS_POSTO_105" := "BYPASS_STATION_105";
   "BYPASS_POSTO_110" := "BYPASS_STATION_110";
   "BYPASS_POSTO_115" := "BYPASS_STATION_115";
   "BYPASS_POSTO_120" := "BYPASS_STATION_120";
   "BYPASS_POSTO_125" := "BYPASS_STATION_125";
   "BYPASS_POSTO_130" := "BYPASS_STATION_130";
   "BYPASS_POSTO_140" := "BYPASS_STATION_140";
   "BYPASS_POSTO_150" := "BYPASS_STATION_150";
   "BYPASS_POSTO_QG" := "BYPASS_STATION_QG";
END_REGION
END_FUNCTION

FUNCTION "Interlock dos sinais linha" : Void   // FC9, LAD
{ S7_Optimized_Access := 'TRUE' }
// stored: SetENOAutomatically false
   VAR_TEMP
      SIGNAL_HELGE : Bool;
      SIGNAL_HELGE1 : Bool;
   END_VAR
   VAR_TEMP   // added for the SCL form of the ladder/FBD networks
      _w1 : Bool;
      _w2 : Bool;
      _w3 : Bool;
      _w4 : Bool;
   END_VAR
BEGIN

REGION Network 1: SCADA DESABILITADO
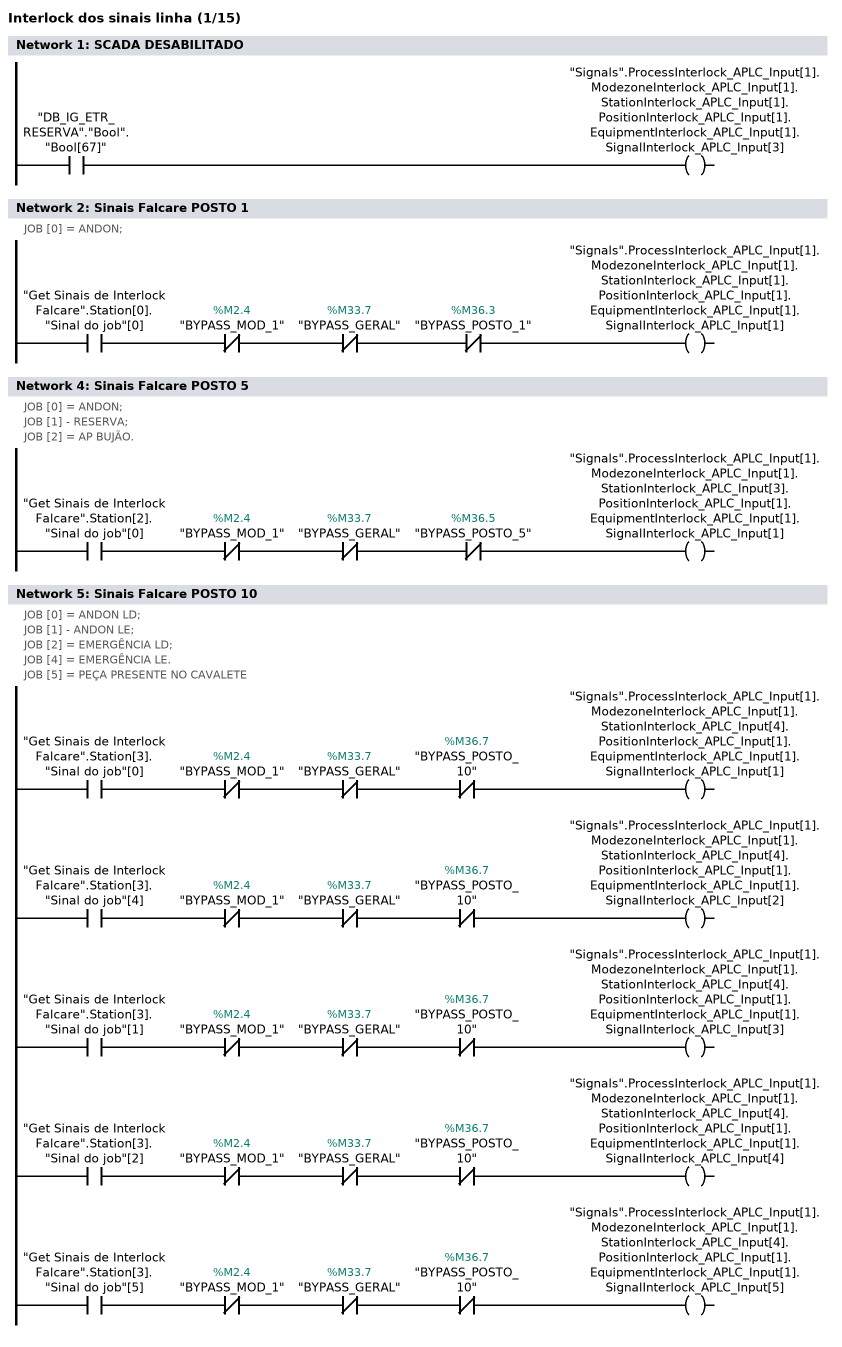
   RUNG wire#powerrail
      Contact( "DB_IG_ETR_RESERVA"."Bool"."Bool[67]" )
      Coil( "Signals".ProcessInterlock_APLC_Input[1].ModezoneInterlock_APLC_Input[1].StationInterlock_APLC_Input[1].PositionInterlock_APLC_Input[1].EquipmentInterlock_APLC_Input[1].SignalInterlock_APLC_Input[3] )
   END_RUNG
   // the same network as SCL:
   "Signals".ProcessInterlock_APLC_Input[1].ModezoneInterlock_APLC_Input[1].StationInterlock_APLC_Input[1].PositionInterlock_APLC_Input[1].EquipmentInterlock_APLC_Input[1].SignalInterlock_APLC_Input[3] := "DB_IG_ETR_RESERVA"."Bool"."Bool[67]";
END_REGION

REGION Network 2: Sinais Falcare POSTO 1
   // JOB [0] = ANDON;
   RUNG wire#powerrail
      Contact( "Get Sinais de Interlock Falcare".Station[0]."Sinal do job"[0] )
      I_Contact( "BYPASS_MOD_1" )
      I_Contact( "BYPASS_GERAL" )
      I_Contact( "BYPASS_POSTO_1" )
      Coil( "Signals".ProcessInterlock_APLC_Input[1].ModezoneInterlock_APLC_Input[1].StationInterlock_APLC_Input[1].PositionInterlock_APLC_Input[1].EquipmentInterlock_APLC_Input[1].SignalInterlock_APLC_Input[1] )
   END_RUNG
   // the same network as SCL:
   "Signals".ProcessInterlock_APLC_Input[1].ModezoneInterlock_APLC_Input[1].StationInterlock_APLC_Input[1].PositionInterlock_APLC_Input[1].EquipmentInterlock_APLC_Input[1].SignalInterlock_APLC_Input[1] := "Get Sinais de Interlock Falcare".Station[0]."Sinal do job"[0] AND NOT "BYPASS_MOD_1" AND NOT "BYPASS_GERAL" AND NOT "BYPASS_POSTO_1";
END_REGION

REGION Network 3: Sinais Falcare VIVERK
   // JOB [0] = ANDON;
   // JOB [1] - EMERGÊNCIA;
END_REGION

REGION Network 4: Sinais Falcare POSTO 5
   // JOB [0] = ANDON;
   // JOB [1] - RESERVA;
   // JOB [2] = AP BUJÃO.
   RUNG wire#powerrail
      Contact( "Get Sinais de Interlock Falcare".Station[2]."Sinal do job"[0] )
      I_Contact( "BYPASS_MOD_1" )
      I_Contact( "BYPASS_GERAL" )
      I_Contact( "BYPASS_POSTO_5" )
      Coil( "Signals".ProcessInterlock_APLC_Input[1].ModezoneInterlock_APLC_Input[1].StationInterlock_APLC_Input[3].PositionInterlock_APLC_Input[1].EquipmentInterlock_APLC_Input[1].SignalInterlock_APLC_Input[1] )
   END_RUNG
   // the same network as SCL:
   "Signals".ProcessInterlock_APLC_Input[1].ModezoneInterlock_APLC_Input[1].StationInterlock_APLC_Input[3].PositionInterlock_APLC_Input[1].EquipmentInterlock_APLC_Input[1].SignalInterlock_APLC_Input[1] := "Get Sinais de Interlock Falcare".Station[2]."Sinal do job"[0] AND NOT "BYPASS_MOD_1" AND NOT "BYPASS_GERAL" AND NOT "BYPASS_POSTO_5";
END_REGION

REGION Network 5: Sinais Falcare POSTO 10
   // JOB [0] = ANDON LD;
   // JOB [1] - ANDON LE;
   // JOB [2] = EMERGÊNCIA LD;
   // JOB [4] = EMERGÊNCIA LE.
   // JOB [5] = PEÇA PRESENTE NO CAVALETE
   RUNG wire#powerrail
      Contact( "Get Sinais de Interlock Falcare".Station[3]."Sinal do job"[0] )
      I_Contact( "BYPASS_MOD_1" )
      I_Contact( "BYPASS_GERAL" )
      I_Contact( "BYPASS_POSTO_10" )
      Coil( "Signals".ProcessInterlock_APLC_Input[1].ModezoneInterlock_APLC_Input[1].StationInterlock_APLC_Input[4].PositionInterlock_APLC_Input[1].EquipmentInterlock_APLC_Input[1].SignalInterlock_APLC_Input[1] )
   END_RUNG
   RUNG wire#powerrail
      Contact( "Get Sinais de Interlock Falcare".Station[3]."Sinal do job"[4] )
      I_Contact( "BYPASS_MOD_1" )
      I_Contact( "BYPASS_GERAL" )
      I_Contact( "BYPASS_POSTO_10" )
      Coil( "Signals".ProcessInterlock_APLC_Input[1].ModezoneInterlock_APLC_Input[1].StationInterlock_APLC_Input[4].PositionInterlock_APLC_Input[1].EquipmentInterlock_APLC_Input[1].SignalInterlock_APLC_Input[2] )
   END_RUNG
   RUNG wire#powerrail
      Contact( "Get Sinais de Interlock Falcare".Station[3]."Sinal do job"[1] )
      I_Contact( "BYPASS_MOD_1" )
      I_Contact( "BYPASS_GERAL" )
      I_Contact( "BYPASS_POSTO_10" )
      Coil( "Signals".ProcessInterlock_APLC_Input[1].ModezoneInterlock_APLC_Input[1].StationInterlock_APLC_Input[4].PositionInterlock_APLC_Input[1].EquipmentInterlock_APLC_Input[1].SignalInterlock_APLC_Input[3] )
   END_RUNG
   RUNG wire#powerrail
      Contact( "Get Sinais de Interlock Falcare".Station[3]."Sinal do job"[2] )
      I_Contact( "BYPASS_MOD_1" )
      I_Contact( "BYPASS_GERAL" )
      I_Contact( "BYPASS_POSTO_10" )
      Coil( "Signals".ProcessInterlock_APLC_Input[1].ModezoneInterlock_APLC_Input[1].StationInterlock_APLC_Input[4].PositionInterlock_APLC_Input[1].EquipmentInterlock_APLC_Input[1].SignalInterlock_APLC_Input[4] )
   END_RUNG
   RUNG wire#powerrail
      Contact( "Get Sinais de Interlock Falcare".Station[3]."Sinal do job"[5] )
      I_Contact( "BYPASS_MOD_1" )
      I_Contact( "BYPASS_GERAL" )
      I_Contact( "BYPASS_POSTO_10" )
      Coil( "Signals".ProcessInterlock_APLC_Input[1].ModezoneInterlock_APLC_Input[1].StationInterlock_APLC_Input[4].PositionInterlock_APLC_Input[1].EquipmentInterlock_APLC_Input[1].SignalInterlock_APLC_Input[5] )
   END_RUNG
   // the same network as SCL:
   "Signals".ProcessInterlock_APLC_Input[1].ModezoneInterlock_APLC_Input[1].StationInterlock_APLC_Input[4].PositionInterlock_APLC_Input[1].EquipmentInterlock_APLC_Input[1].SignalInterlock_APLC_Input[1] := "Get Sinais de Interlock Falcare".Station[3]."Sinal do job"[0] AND NOT "BYPASS_MOD_1" AND NOT "BYPASS_GERAL" AND NOT "BYPASS_POSTO_10";
   "Signals".ProcessInterlock_APLC_Input[1].ModezoneInterlock_APLC_Input[1].StationInterlock_APLC_Input[4].PositionInterlock_APLC_Input[1].EquipmentInterlock_APLC_Input[1].SignalInterlock_APLC_Input[2] := "Get Sinais de Interlock Falcare".Station[3]."Sinal do job"[4] AND NOT "BYPASS_MOD_1" AND NOT "BYPASS_GERAL" AND NOT "BYPASS_POSTO_10";
   "Signals".ProcessInterlock_APLC_Input[1].ModezoneInterlock_APLC_Input[1].StationInterlock_APLC_Input[4].PositionInterlock_APLC_Input[1].EquipmentInterlock_APLC_Input[1].SignalInterlock_APLC_Input[3] := "Get Sinais de Interlock Falcare".Station[3]."Sinal do job"[1] AND NOT "BYPASS_MOD_1" AND NOT "BYPASS_GERAL" AND NOT "BYPASS_POSTO_10";
   "Signals".ProcessInterlock_APLC_Input[1].ModezoneInterlock_APLC_Input[1].StationInterlock_APLC_Input[4].PositionInterlock_APLC_Input[1].EquipmentInterlock_APLC_Input[1].SignalInterlock_APLC_Input[4] := "Get Sinais de Interlock Falcare".Station[3]."Sinal do job"[2] AND NOT "BYPASS_MOD_1" AND NOT "BYPASS_GERAL" AND NOT "BYPASS_POSTO_10";
   "Signals".ProcessInterlock_APLC_Input[1].ModezoneInterlock_APLC_Input[1].StationInterlock_APLC_Input[4].PositionInterlock_APLC_Input[1].EquipmentInterlock_APLC_Input[1].SignalInterlock_APLC_Input[5] := "Get Sinais de Interlock Falcare".Station[3]."Sinal do job"[5] AND NOT "BYPASS_MOD_1" AND NOT "BYPASS_GERAL" AND NOT "BYPASS_POSTO_10";
END_REGION

REGION Network 6: Sinais Falcare POSTO 15
   // JOB [3] = AP TUBO RPX POSTO 15;
END_REGION

REGION Network 7: Sinais Falcare POSTO 20
   // JOB [0] = ANDON LD;
   // JOB [1] - EMERGÊNCIA LD;
   // JOB [2] = AP MOLA HARPA;
   // JOB [3] = SENSOR POSIÇÃO AP HARPA;
   // JOB [4] = AP TUBO LUBRIFICAÇÃO RPX I9.0
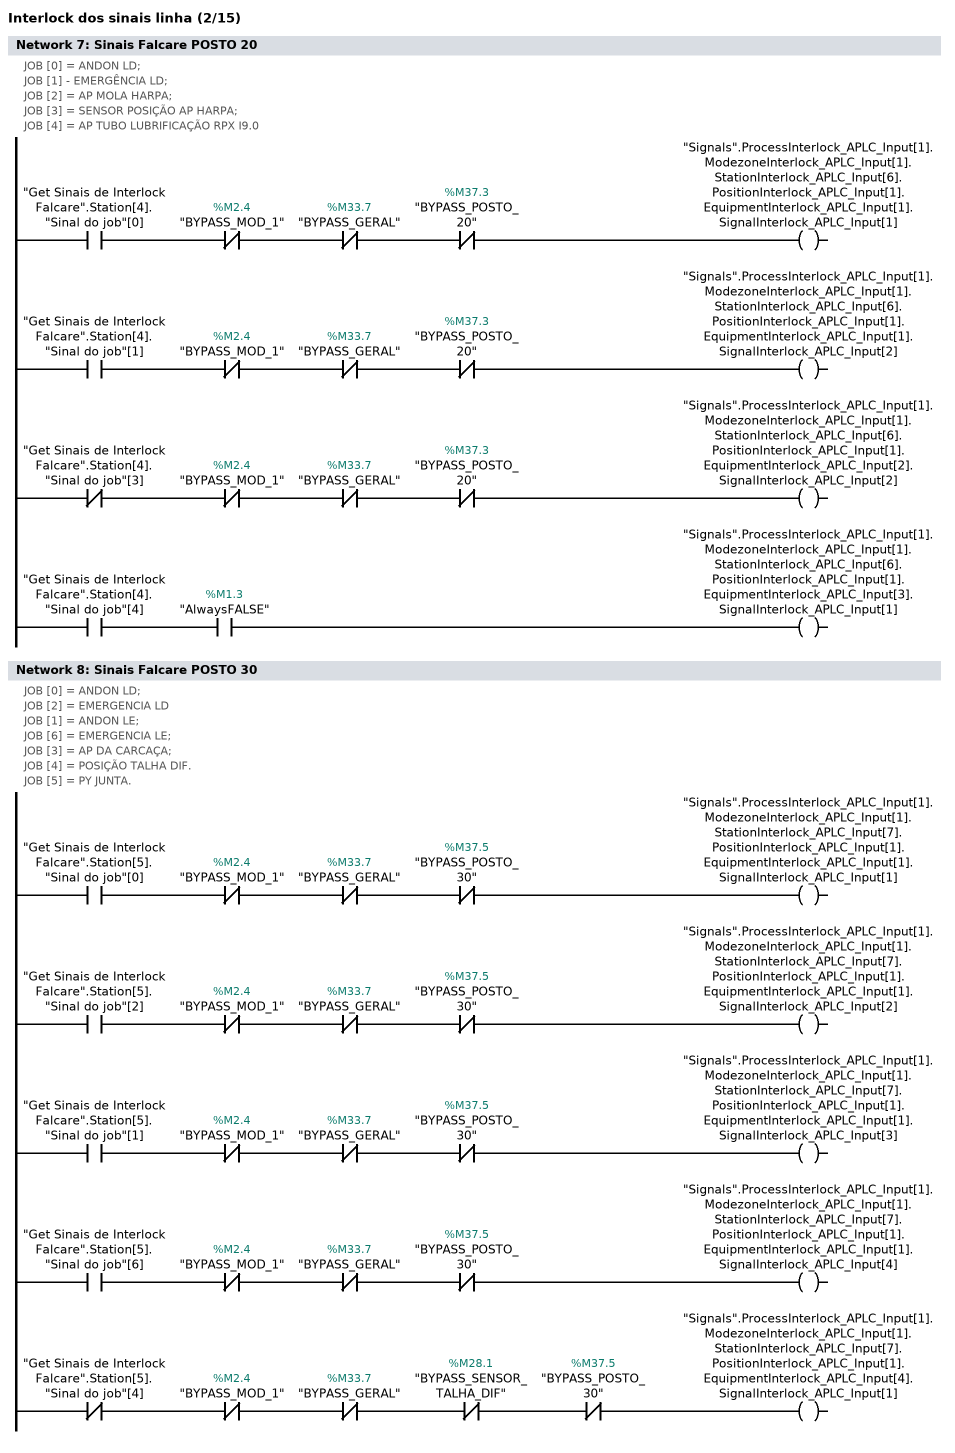
   RUNG wire#powerrail
      Contact( "Get Sinais de Interlock Falcare".Station[4]."Sinal do job"[0] )
      I_Contact( "BYPASS_MOD_1" )
      I_Contact( "BYPASS_GERAL" )
      I_Contact( "BYPASS_POSTO_20" )
      Coil( "Signals".ProcessInterlock_APLC_Input[1].ModezoneInterlock_APLC_Input[1].StationInterlock_APLC_Input[6].PositionInterlock_APLC_Input[1].EquipmentInterlock_APLC_Input[1].SignalInterlock_APLC_Input[1] )
   END_RUNG
   RUNG wire#powerrail
      Contact( "Get Sinais de Interlock Falcare".Station[4]."Sinal do job"[1] )
      I_Contact( "BYPASS_MOD_1" )
      I_Contact( "BYPASS_GERAL" )
      I_Contact( "BYPASS_POSTO_20" )
      Coil( "Signals".ProcessInterlock_APLC_Input[1].ModezoneInterlock_APLC_Input[1].StationInterlock_APLC_Input[6].PositionInterlock_APLC_Input[1].EquipmentInterlock_APLC_Input[1].SignalInterlock_APLC_Input[2] )
   END_RUNG
   RUNG wire#powerrail
      I_Contact( "Get Sinais de Interlock Falcare".Station[4]."Sinal do job"[3] )
      I_Contact( "BYPASS_MOD_1" )
      I_Contact( "BYPASS_GERAL" )
      I_Contact( "BYPASS_POSTO_20" )
      Coil( "Signals".ProcessInterlock_APLC_Input[1].ModezoneInterlock_APLC_Input[1].StationInterlock_APLC_Input[6].PositionInterlock_APLC_Input[1].EquipmentInterlock_APLC_Input[2].SignalInterlock_APLC_Input[2] )
   END_RUNG
   RUNG wire#powerrail
      Contact( "Get Sinais de Interlock Falcare".Station[4]."Sinal do job"[4] )
      Contact( "AlwaysFALSE" )
      Coil( "Signals".ProcessInterlock_APLC_Input[1].ModezoneInterlock_APLC_Input[1].StationInterlock_APLC_Input[6].PositionInterlock_APLC_Input[1].EquipmentInterlock_APLC_Input[3].SignalInterlock_APLC_Input[1] )
   END_RUNG
   // the same network as SCL:
   "Signals".ProcessInterlock_APLC_Input[1].ModezoneInterlock_APLC_Input[1].StationInterlock_APLC_Input[6].PositionInterlock_APLC_Input[1].EquipmentInterlock_APLC_Input[1].SignalInterlock_APLC_Input[1] := "Get Sinais de Interlock Falcare".Station[4]."Sinal do job"[0] AND NOT "BYPASS_MOD_1" AND NOT "BYPASS_GERAL" AND NOT "BYPASS_POSTO_20";
   "Signals".ProcessInterlock_APLC_Input[1].ModezoneInterlock_APLC_Input[1].StationInterlock_APLC_Input[6].PositionInterlock_APLC_Input[1].EquipmentInterlock_APLC_Input[1].SignalInterlock_APLC_Input[2] := "Get Sinais de Interlock Falcare".Station[4]."Sinal do job"[1] AND NOT "BYPASS_MOD_1" AND NOT "BYPASS_GERAL" AND NOT "BYPASS_POSTO_20";
   "Signals".ProcessInterlock_APLC_Input[1].ModezoneInterlock_APLC_Input[1].StationInterlock_APLC_Input[6].PositionInterlock_APLC_Input[1].EquipmentInterlock_APLC_Input[2].SignalInterlock_APLC_Input[2] := NOT "Get Sinais de Interlock Falcare".Station[4]."Sinal do job"[3] AND NOT "BYPASS_MOD_1" AND NOT "BYPASS_GERAL" AND NOT "BYPASS_POSTO_20";
   "Signals".ProcessInterlock_APLC_Input[1].ModezoneInterlock_APLC_Input[1].StationInterlock_APLC_Input[6].PositionInterlock_APLC_Input[1].EquipmentInterlock_APLC_Input[3].SignalInterlock_APLC_Input[1] := "Get Sinais de Interlock Falcare".Station[4]."Sinal do job"[4] AND "AlwaysFALSE";
END_REGION

REGION Network 8: Sinais Falcare POSTO 30
   // JOB [0] = ANDON LD;
   // JOB [2] = EMERGENCIA LD
   // JOB [1] = ANDON LE;
   // JOB [6] = EMERGENCIA LE;
   // JOB [3] = AP DA CARCAÇA;
   // JOB [4] = POSIÇÃO TALHA DIF.
   // JOB [5] = PY JUNTA.
   RUNG wire#powerrail
      Contact( "Get Sinais de Interlock Falcare".Station[5]."Sinal do job"[0] )
      I_Contact( "BYPASS_MOD_1" )
      I_Contact( "BYPASS_GERAL" )
      I_Contact( "BYPASS_POSTO_30" )
      Coil( "Signals".ProcessInterlock_APLC_Input[1].ModezoneInterlock_APLC_Input[1].StationInterlock_APLC_Input[7].PositionInterlock_APLC_Input[1].EquipmentInterlock_APLC_Input[1].SignalInterlock_APLC_Input[1] )
   END_RUNG
   RUNG wire#powerrail
      Contact( "Get Sinais de Interlock Falcare".Station[5]."Sinal do job"[2] )
      I_Contact( "BYPASS_MOD_1" )
      I_Contact( "BYPASS_GERAL" )
      I_Contact( "BYPASS_POSTO_30" )
      Coil( "Signals".ProcessInterlock_APLC_Input[1].ModezoneInterlock_APLC_Input[1].StationInterlock_APLC_Input[7].PositionInterlock_APLC_Input[1].EquipmentInterlock_APLC_Input[1].SignalInterlock_APLC_Input[2] )
   END_RUNG
   RUNG wire#powerrail
      Contact( "Get Sinais de Interlock Falcare".Station[5]."Sinal do job"[1] )
      I_Contact( "BYPASS_MOD_1" )
      I_Contact( "BYPASS_GERAL" )
      I_Contact( "BYPASS_POSTO_30" )
      Coil( "Signals".ProcessInterlock_APLC_Input[1].ModezoneInterlock_APLC_Input[1].StationInterlock_APLC_Input[7].PositionInterlock_APLC_Input[1].EquipmentInterlock_APLC_Input[1].SignalInterlock_APLC_Input[3] )
   END_RUNG
   RUNG wire#powerrail
      Contact( "Get Sinais de Interlock Falcare".Station[5]."Sinal do job"[6] )
      I_Contact( "BYPASS_MOD_1" )
      I_Contact( "BYPASS_GERAL" )
      I_Contact( "BYPASS_POSTO_30" )
      Coil( "Signals".ProcessInterlock_APLC_Input[1].ModezoneInterlock_APLC_Input[1].StationInterlock_APLC_Input[7].PositionInterlock_APLC_Input[1].EquipmentInterlock_APLC_Input[1].SignalInterlock_APLC_Input[4] )
   END_RUNG
   RUNG wire#powerrail
      I_Contact( "Get Sinais de Interlock Falcare".Station[5]."Sinal do job"[4] )
      I_Contact( "BYPASS_MOD_1" )
      I_Contact( "BYPASS_GERAL" )
      I_Contact( "BYPASS_SENSOR_TALHA_DIF" )
      I_Contact( "BYPASS_POSTO_30" )
      Coil( "Signals".ProcessInterlock_APLC_Input[1].ModezoneInterlock_APLC_Input[1].StationInterlock_APLC_Input[7].PositionInterlock_APLC_Input[1].EquipmentInterlock_APLC_Input[4].SignalInterlock_APLC_Input[1] )
   END_RUNG
   // the same network as SCL:
   "Signals".ProcessInterlock_APLC_Input[1].ModezoneInterlock_APLC_Input[1].StationInterlock_APLC_Input[7].PositionInterlock_APLC_Input[1].EquipmentInterlock_APLC_Input[1].SignalInterlock_APLC_Input[1] := "Get Sinais de Interlock Falcare".Station[5]."Sinal do job"[0] AND NOT "BYPASS_MOD_1" AND NOT "BYPASS_GERAL" AND NOT "BYPASS_POSTO_30";
   "Signals".ProcessInterlock_APLC_Input[1].ModezoneInterlock_APLC_Input[1].StationInterlock_APLC_Input[7].PositionInterlock_APLC_Input[1].EquipmentInterlock_APLC_Input[1].SignalInterlock_APLC_Input[2] := "Get Sinais de Interlock Falcare".Station[5]."Sinal do job"[2] AND NOT "BYPASS_MOD_1" AND NOT "BYPASS_GERAL" AND NOT "BYPASS_POSTO_30";
   "Signals".ProcessInterlock_APLC_Input[1].ModezoneInterlock_APLC_Input[1].StationInterlock_APLC_Input[7].PositionInterlock_APLC_Input[1].EquipmentInterlock_APLC_Input[1].SignalInterlock_APLC_Input[3] := "Get Sinais de Interlock Falcare".Station[5]."Sinal do job"[1] AND NOT "BYPASS_MOD_1" AND NOT "BYPASS_GERAL" AND NOT "BYPASS_POSTO_30";
   "Signals".ProcessInterlock_APLC_Input[1].ModezoneInterlock_APLC_Input[1].StationInterlock_APLC_Input[7].PositionInterlock_APLC_Input[1].EquipmentInterlock_APLC_Input[1].SignalInterlock_APLC_Input[4] := "Get Sinais de Interlock Falcare".Station[5]."Sinal do job"[6] AND NOT "BYPASS_MOD_1" AND NOT "BYPASS_GERAL" AND NOT "BYPASS_POSTO_30";
   "Signals".ProcessInterlock_APLC_Input[1].ModezoneInterlock_APLC_Input[1].StationInterlock_APLC_Input[7].PositionInterlock_APLC_Input[1].EquipmentInterlock_APLC_Input[4].SignalInterlock_APLC_Input[1] := NOT "Get Sinais de Interlock Falcare".Station[5]."Sinal do job"[4] AND NOT "BYPASS_MOD_1" AND NOT "BYPASS_GERAL" AND NOT "BYPASS_SENSOR_TALHA_DIF" AND NOT "BYPASS_POSTO_30";
END_REGION

REGION Network 9: Sinais Falcare POSTO 40
   // JOB [0] = ANDON LD;
   // JOB [1] = ANDON LE;
   // JOB [2] = EMERGENCIA LE;
   // JOB [3] = AP CRAWFOOT PORCA;
   // JOB [4] = SENSOR POSIÇÃO AP CRAWFOOT;
   // JOB [5] = AP PORCA DUPLO FUSO;
   // JOB [6] = SENSOR POSIÇÃO AP DUPLO FUSO;
   // JOB [7] = EMERGÊNCIA LD.
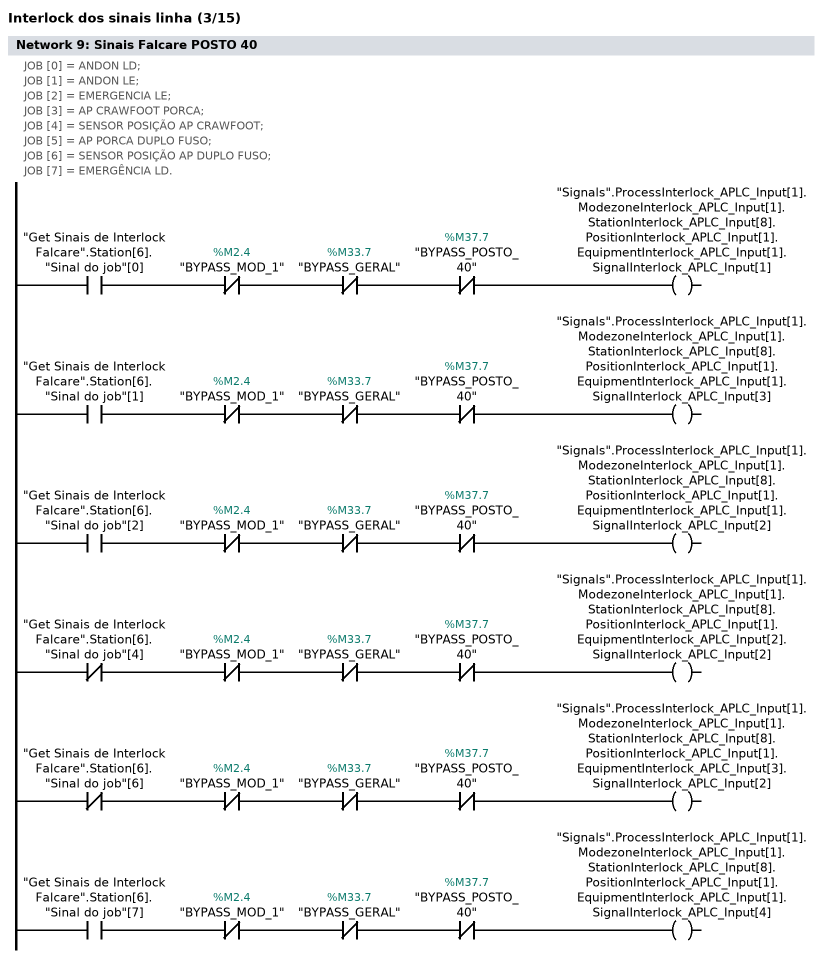
   RUNG wire#powerrail
      Contact( "Get Sinais de Interlock Falcare".Station[6]."Sinal do job"[0] )
      I_Contact( "BYPASS_MOD_1" )
      I_Contact( "BYPASS_GERAL" )
      I_Contact( "BYPASS_POSTO_40" )
      Coil( "Signals".ProcessInterlock_APLC_Input[1].ModezoneInterlock_APLC_Input[1].StationInterlock_APLC_Input[8].PositionInterlock_APLC_Input[1].EquipmentInterlock_APLC_Input[1].SignalInterlock_APLC_Input[1] )
   END_RUNG
   RUNG wire#powerrail
      Contact( "Get Sinais de Interlock Falcare".Station[6]."Sinal do job"[1] )
      I_Contact( "BYPASS_MOD_1" )
      I_Contact( "BYPASS_GERAL" )
      I_Contact( "BYPASS_POSTO_40" )
      Coil( "Signals".ProcessInterlock_APLC_Input[1].ModezoneInterlock_APLC_Input[1].StationInterlock_APLC_Input[8].PositionInterlock_APLC_Input[1].EquipmentInterlock_APLC_Input[1].SignalInterlock_APLC_Input[3] )
   END_RUNG
   RUNG wire#powerrail
      Contact( "Get Sinais de Interlock Falcare".Station[6]."Sinal do job"[2] )
      I_Contact( "BYPASS_MOD_1" )
      I_Contact( "BYPASS_GERAL" )
      I_Contact( "BYPASS_POSTO_40" )
      Coil( "Signals".ProcessInterlock_APLC_Input[1].ModezoneInterlock_APLC_Input[1].StationInterlock_APLC_Input[8].PositionInterlock_APLC_Input[1].EquipmentInterlock_APLC_Input[1].SignalInterlock_APLC_Input[2] )
   END_RUNG
   RUNG wire#powerrail
      I_Contact( "Get Sinais de Interlock Falcare".Station[6]."Sinal do job"[4] )
      I_Contact( "BYPASS_MOD_1" )
      I_Contact( "BYPASS_GERAL" )
      I_Contact( "BYPASS_POSTO_40" )
      Coil( "Signals".ProcessInterlock_APLC_Input[1].ModezoneInterlock_APLC_Input[1].StationInterlock_APLC_Input[8].PositionInterlock_APLC_Input[1].EquipmentInterlock_APLC_Input[2].SignalInterlock_APLC_Input[2] )
   END_RUNG
   RUNG wire#powerrail
      I_Contact( "Get Sinais de Interlock Falcare".Station[6]."Sinal do job"[6] )
      I_Contact( "BYPASS_MOD_1" )
      I_Contact( "BYPASS_GERAL" )
      I_Contact( "BYPASS_POSTO_40" )
      Coil( "Signals".ProcessInterlock_APLC_Input[1].ModezoneInterlock_APLC_Input[1].StationInterlock_APLC_Input[8].PositionInterlock_APLC_Input[1].EquipmentInterlock_APLC_Input[3].SignalInterlock_APLC_Input[2] )
   END_RUNG
   RUNG wire#powerrail
      Contact( "Get Sinais de Interlock Falcare".Station[6]."Sinal do job"[7] )
      I_Contact( "BYPASS_MOD_1" )
      I_Contact( "BYPASS_GERAL" )
      I_Contact( "BYPASS_POSTO_40" )
      Coil( "Signals".ProcessInterlock_APLC_Input[1].ModezoneInterlock_APLC_Input[1].StationInterlock_APLC_Input[8].PositionInterlock_APLC_Input[1].EquipmentInterlock_APLC_Input[1].SignalInterlock_APLC_Input[4] )
   END_RUNG
   // the same network as SCL:
   "Signals".ProcessInterlock_APLC_Input[1].ModezoneInterlock_APLC_Input[1].StationInterlock_APLC_Input[8].PositionInterlock_APLC_Input[1].EquipmentInterlock_APLC_Input[1].SignalInterlock_APLC_Input[1] := "Get Sinais de Interlock Falcare".Station[6]."Sinal do job"[0] AND NOT "BYPASS_MOD_1" AND NOT "BYPASS_GERAL" AND NOT "BYPASS_POSTO_40";
   "Signals".ProcessInterlock_APLC_Input[1].ModezoneInterlock_APLC_Input[1].StationInterlock_APLC_Input[8].PositionInterlock_APLC_Input[1].EquipmentInterlock_APLC_Input[1].SignalInterlock_APLC_Input[3] := "Get Sinais de Interlock Falcare".Station[6]."Sinal do job"[1] AND NOT "BYPASS_MOD_1" AND NOT "BYPASS_GERAL" AND NOT "BYPASS_POSTO_40";
   "Signals".ProcessInterlock_APLC_Input[1].ModezoneInterlock_APLC_Input[1].StationInterlock_APLC_Input[8].PositionInterlock_APLC_Input[1].EquipmentInterlock_APLC_Input[1].SignalInterlock_APLC_Input[2] := "Get Sinais de Interlock Falcare".Station[6]."Sinal do job"[2] AND NOT "BYPASS_MOD_1" AND NOT "BYPASS_GERAL" AND NOT "BYPASS_POSTO_40";
   "Signals".ProcessInterlock_APLC_Input[1].ModezoneInterlock_APLC_Input[1].StationInterlock_APLC_Input[8].PositionInterlock_APLC_Input[1].EquipmentInterlock_APLC_Input[2].SignalInterlock_APLC_Input[2] := NOT "Get Sinais de Interlock Falcare".Station[6]."Sinal do job"[4] AND NOT "BYPASS_MOD_1" AND NOT "BYPASS_GERAL" AND NOT "BYPASS_POSTO_40";
   "Signals".ProcessInterlock_APLC_Input[1].ModezoneInterlock_APLC_Input[1].StationInterlock_APLC_Input[8].PositionInterlock_APLC_Input[1].EquipmentInterlock_APLC_Input[3].SignalInterlock_APLC_Input[2] := NOT "Get Sinais de Interlock Falcare".Station[6]."Sinal do job"[6] AND NOT "BYPASS_MOD_1" AND NOT "BYPASS_GERAL" AND NOT "BYPASS_POSTO_40";
   "Signals".ProcessInterlock_APLC_Input[1].ModezoneInterlock_APLC_Input[1].StationInterlock_APLC_Input[8].PositionInterlock_APLC_Input[1].EquipmentInterlock_APLC_Input[1].SignalInterlock_APLC_Input[4] := "Get Sinais de Interlock Falcare".Station[6]."Sinal do job"[7] AND NOT "BYPASS_MOD_1" AND NOT "BYPASS_GERAL" AND NOT "BYPASS_POSTO_40";
END_REGION

REGION Network 10: Sinais Falcare POSTO 50
   // JOB [0] = ANDON;
   // JOB [1] = EMERGENCIA;
   // JOB [2] = AP PORCA ESCONDIDA;
   // JOB [3] = SENSOR POSIÇÃO AP PORCA ESCONDIDA;
   // JOB [4] = AP PORCA SUPORTE DO CILINDRO;
   // JOB [5] = SENSOR POSIÇÃO AP SUPORTE DO CILINDRO;
   // JOB [7] = AP VÁLVULA
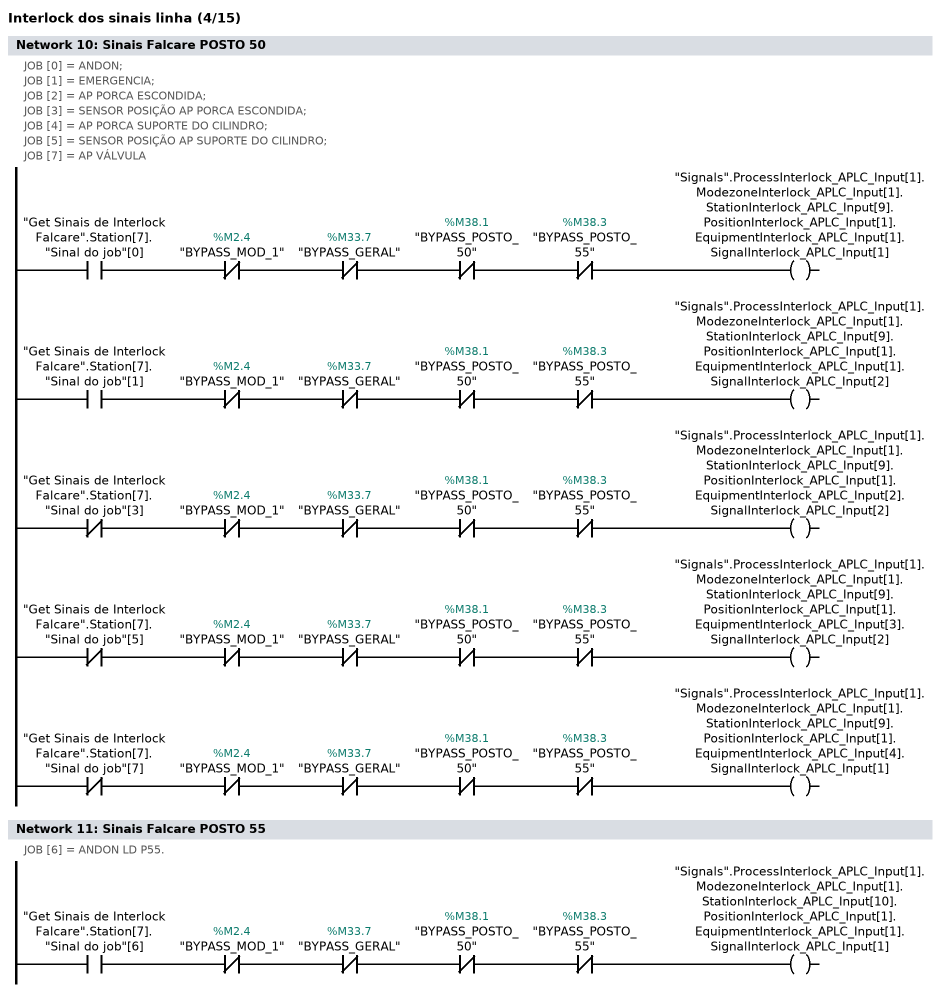
   RUNG wire#powerrail
      Contact( "Get Sinais de Interlock Falcare".Station[7]."Sinal do job"[0] )
      I_Contact( "BYPASS_MOD_1" )
      I_Contact( "BYPASS_GERAL" )
      I_Contact( "BYPASS_POSTO_50" )
      I_Contact( "BYPASS_POSTO_55" )
      Coil( "Signals".ProcessInterlock_APLC_Input[1].ModezoneInterlock_APLC_Input[1].StationInterlock_APLC_Input[9].PositionInterlock_APLC_Input[1].EquipmentInterlock_APLC_Input[1].SignalInterlock_APLC_Input[1] )
   END_RUNG
   RUNG wire#powerrail
      Contact( "Get Sinais de Interlock Falcare".Station[7]."Sinal do job"[1] )
      I_Contact( "BYPASS_MOD_1" )
      I_Contact( "BYPASS_GERAL" )
      I_Contact( "BYPASS_POSTO_50" )
      I_Contact( "BYPASS_POSTO_55" )
      Coil( "Signals".ProcessInterlock_APLC_Input[1].ModezoneInterlock_APLC_Input[1].StationInterlock_APLC_Input[9].PositionInterlock_APLC_Input[1].EquipmentInterlock_APLC_Input[1].SignalInterlock_APLC_Input[2] )
   END_RUNG
   RUNG wire#powerrail
      I_Contact( "Get Sinais de Interlock Falcare".Station[7]."Sinal do job"[3] )
      I_Contact( "BYPASS_MOD_1" )
      I_Contact( "BYPASS_GERAL" )
      I_Contact( "BYPASS_POSTO_50" )
      I_Contact( "BYPASS_POSTO_55" )
      Coil( "Signals".ProcessInterlock_APLC_Input[1].ModezoneInterlock_APLC_Input[1].StationInterlock_APLC_Input[9].PositionInterlock_APLC_Input[1].EquipmentInterlock_APLC_Input[2].SignalInterlock_APLC_Input[2] )
   END_RUNG
   RUNG wire#powerrail
      I_Contact( "Get Sinais de Interlock Falcare".Station[7]."Sinal do job"[5] )
      I_Contact( "BYPASS_MOD_1" )
      I_Contact( "BYPASS_GERAL" )
      I_Contact( "BYPASS_POSTO_50" )
      I_Contact( "BYPASS_POSTO_55" )
      Coil( "Signals".ProcessInterlock_APLC_Input[1].ModezoneInterlock_APLC_Input[1].StationInterlock_APLC_Input[9].PositionInterlock_APLC_Input[1].EquipmentInterlock_APLC_Input[3].SignalInterlock_APLC_Input[2] )
   END_RUNG
   RUNG wire#powerrail
      I_Contact( "Get Sinais de Interlock Falcare".Station[7]."Sinal do job"[7] )
      I_Contact( "BYPASS_MOD_1" )
      I_Contact( "BYPASS_GERAL" )
      I_Contact( "BYPASS_POSTO_50" )
      I_Contact( "BYPASS_POSTO_55" )
      Coil( "Signals".ProcessInterlock_APLC_Input[1].ModezoneInterlock_APLC_Input[1].StationInterlock_APLC_Input[9].PositionInterlock_APLC_Input[1].EquipmentInterlock_APLC_Input[4].SignalInterlock_APLC_Input[1] )
   END_RUNG
   // the same network as SCL:
   "Signals".ProcessInterlock_APLC_Input[1].ModezoneInterlock_APLC_Input[1].StationInterlock_APLC_Input[9].PositionInterlock_APLC_Input[1].EquipmentInterlock_APLC_Input[1].SignalInterlock_APLC_Input[1] := "Get Sinais de Interlock Falcare".Station[7]."Sinal do job"[0] AND NOT "BYPASS_MOD_1" AND NOT "BYPASS_GERAL" AND NOT "BYPASS_POSTO_50" AND NOT "BYPASS_POSTO_55";
   "Signals".ProcessInterlock_APLC_Input[1].ModezoneInterlock_APLC_Input[1].StationInterlock_APLC_Input[9].PositionInterlock_APLC_Input[1].EquipmentInterlock_APLC_Input[1].SignalInterlock_APLC_Input[2] := "Get Sinais de Interlock Falcare".Station[7]."Sinal do job"[1] AND NOT "BYPASS_MOD_1" AND NOT "BYPASS_GERAL" AND NOT "BYPASS_POSTO_50" AND NOT "BYPASS_POSTO_55";
   "Signals".ProcessInterlock_APLC_Input[1].ModezoneInterlock_APLC_Input[1].StationInterlock_APLC_Input[9].PositionInterlock_APLC_Input[1].EquipmentInterlock_APLC_Input[2].SignalInterlock_APLC_Input[2] := NOT "Get Sinais de Interlock Falcare".Station[7]."Sinal do job"[3] AND NOT "BYPASS_MOD_1" AND NOT "BYPASS_GERAL" AND NOT "BYPASS_POSTO_50" AND NOT "BYPASS_POSTO_55";
   "Signals".ProcessInterlock_APLC_Input[1].ModezoneInterlock_APLC_Input[1].StationInterlock_APLC_Input[9].PositionInterlock_APLC_Input[1].EquipmentInterlock_APLC_Input[3].SignalInterlock_APLC_Input[2] := NOT "Get Sinais de Interlock Falcare".Station[7]."Sinal do job"[5] AND NOT "BYPASS_MOD_1" AND NOT "BYPASS_GERAL" AND NOT "BYPASS_POSTO_50" AND NOT "BYPASS_POSTO_55";
   "Signals".ProcessInterlock_APLC_Input[1].ModezoneInterlock_APLC_Input[1].StationInterlock_APLC_Input[9].PositionInterlock_APLC_Input[1].EquipmentInterlock_APLC_Input[4].SignalInterlock_APLC_Input[1] := NOT "Get Sinais de Interlock Falcare".Station[7]."Sinal do job"[7] AND NOT "BYPASS_MOD_1" AND NOT "BYPASS_GERAL" AND NOT "BYPASS_POSTO_50" AND NOT "BYPASS_POSTO_55";
END_REGION

REGION Network 11: Sinais Falcare POSTO 55
   // JOB [6] = ANDON LD P55.
   RUNG wire#powerrail
      Contact( "Get Sinais de Interlock Falcare".Station[7]."Sinal do job"[6] )
      I_Contact( "BYPASS_MOD_1" )
      I_Contact( "BYPASS_GERAL" )
      I_Contact( "BYPASS_POSTO_50" )
      I_Contact( "BYPASS_POSTO_55" )
      Coil( "Signals".ProcessInterlock_APLC_Input[1].ModezoneInterlock_APLC_Input[1].StationInterlock_APLC_Input[10].PositionInterlock_APLC_Input[1].EquipmentInterlock_APLC_Input[1].SignalInterlock_APLC_Input[1] )
   END_RUNG
   // the same network as SCL:
   "Signals".ProcessInterlock_APLC_Input[1].ModezoneInterlock_APLC_Input[1].StationInterlock_APLC_Input[10].PositionInterlock_APLC_Input[1].EquipmentInterlock_APLC_Input[1].SignalInterlock_APLC_Input[1] := "Get Sinais de Interlock Falcare".Station[7]."Sinal do job"[6] AND NOT "BYPASS_MOD_1" AND NOT "BYPASS_GERAL" AND NOT "BYPASS_POSTO_50" AND NOT "BYPASS_POSTO_55";
END_REGION

REGION Network 12: Sinais Falcare POSTO 60
   // JOB [0] = ANDON;
   // JOB [1] = EMERGENCIA;
   // JOB [2] = AP PORCA DO CILINDRO;
   // JOB [3] = SENSOR POSIÇÃO AP PORCA DO CILINDRO;
   // JOB [4] = EMERGENCIA PAINEL FALCARE.
   // JOB [5] = CONFIRMA PRE AVISO DO GIRADOR
   // JOB [6] = PRODUTO PRESENTE NO GIRADOR (MENSAGEM DE RETIRAR PRODUTO)
   // JOB [7] = FALCARE EM MANUAL
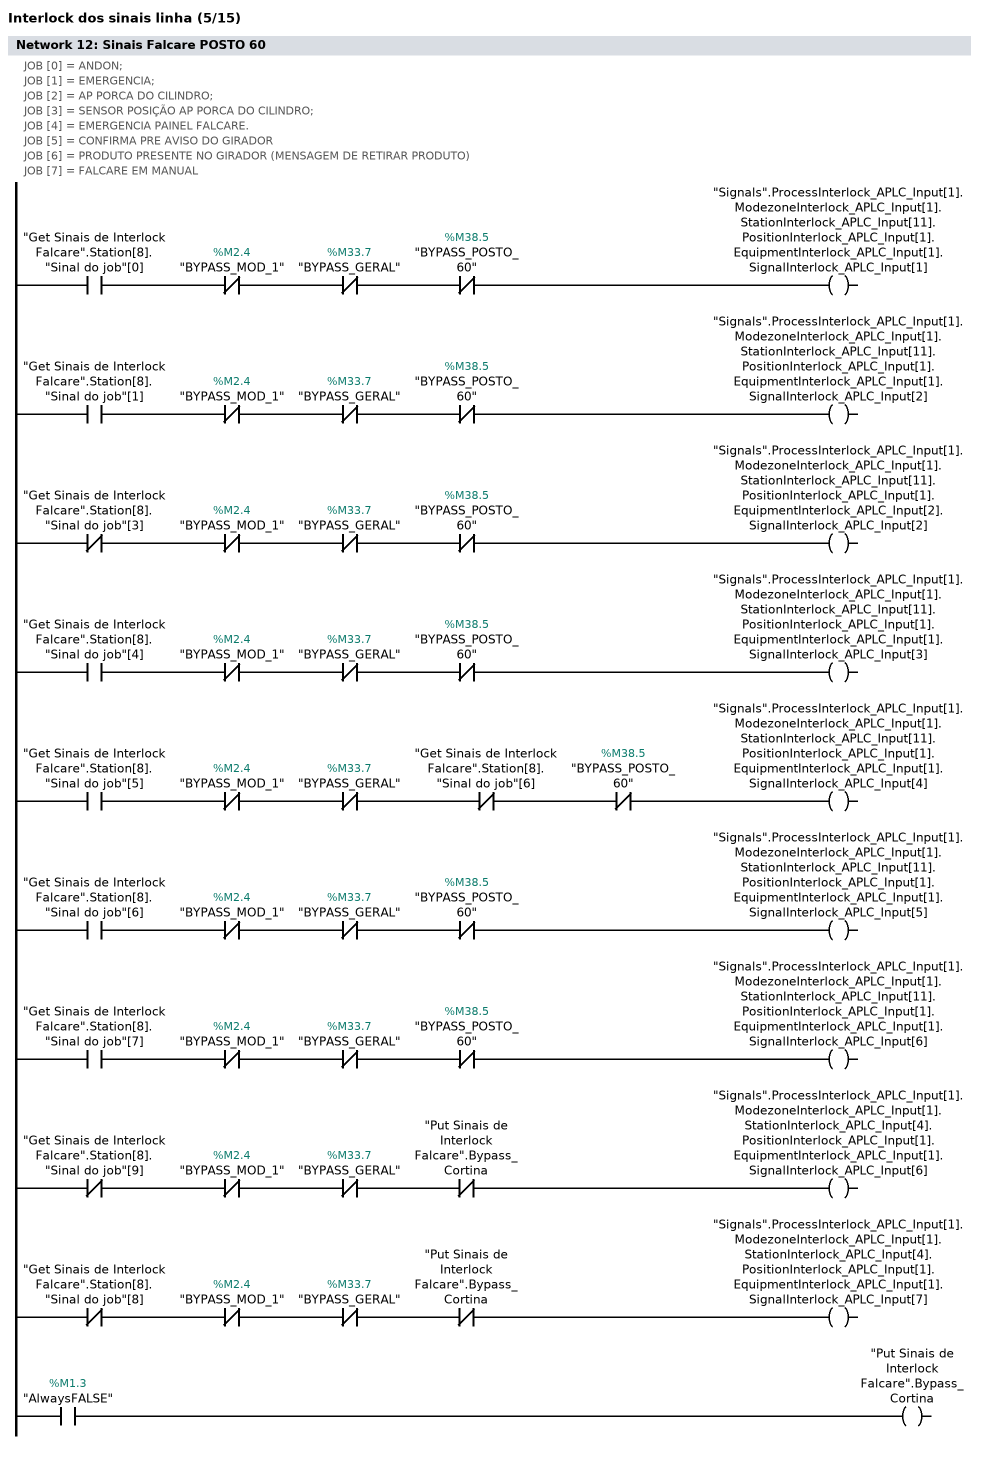
   RUNG wire#powerrail
      Contact( "Get Sinais de Interlock Falcare".Station[8]."Sinal do job"[0] )
      I_Contact( "BYPASS_MOD_1" )
      I_Contact( "BYPASS_GERAL" )
      I_Contact( "BYPASS_POSTO_60" )
      Coil( "Signals".ProcessInterlock_APLC_Input[1].ModezoneInterlock_APLC_Input[1].StationInterlock_APLC_Input[11].PositionInterlock_APLC_Input[1].EquipmentInterlock_APLC_Input[1].SignalInterlock_APLC_Input[1] )
   END_RUNG
   RUNG wire#powerrail
      Contact( "Get Sinais de Interlock Falcare".Station[8]."Sinal do job"[1] )
      I_Contact( "BYPASS_MOD_1" )
      I_Contact( "BYPASS_GERAL" )
      I_Contact( "BYPASS_POSTO_60" )
      Coil( "Signals".ProcessInterlock_APLC_Input[1].ModezoneInterlock_APLC_Input[1].StationInterlock_APLC_Input[11].PositionInterlock_APLC_Input[1].EquipmentInterlock_APLC_Input[1].SignalInterlock_APLC_Input[2] )
   END_RUNG
   RUNG wire#powerrail
      I_Contact( "Get Sinais de Interlock Falcare".Station[8]."Sinal do job"[3] )
      I_Contact( "BYPASS_MOD_1" )
      I_Contact( "BYPASS_GERAL" )
      I_Contact( "BYPASS_POSTO_60" )
      Coil( "Signals".ProcessInterlock_APLC_Input[1].ModezoneInterlock_APLC_Input[1].StationInterlock_APLC_Input[11].PositionInterlock_APLC_Input[1].EquipmentInterlock_APLC_Input[2].SignalInterlock_APLC_Input[2] )
   END_RUNG
   RUNG wire#powerrail
      Contact( "Get Sinais de Interlock Falcare".Station[8]."Sinal do job"[4] )
      I_Contact( "BYPASS_MOD_1" )
      I_Contact( "BYPASS_GERAL" )
      I_Contact( "BYPASS_POSTO_60" )
      Coil( "Signals".ProcessInterlock_APLC_Input[1].ModezoneInterlock_APLC_Input[1].StationInterlock_APLC_Input[11].PositionInterlock_APLC_Input[1].EquipmentInterlock_APLC_Input[1].SignalInterlock_APLC_Input[3] )
   END_RUNG
   RUNG wire#powerrail
      Contact( "Get Sinais de Interlock Falcare".Station[8]."Sinal do job"[5] )
      I_Contact( "BYPASS_MOD_1" )
      I_Contact( "BYPASS_GERAL" )
      I_Contact( "Get Sinais de Interlock Falcare".Station[8]."Sinal do job"[6] )
      I_Contact( "BYPASS_POSTO_60" )
      Coil( "Signals".ProcessInterlock_APLC_Input[1].ModezoneInterlock_APLC_Input[1].StationInterlock_APLC_Input[11].PositionInterlock_APLC_Input[1].EquipmentInterlock_APLC_Input[1].SignalInterlock_APLC_Input[4] )
   END_RUNG
   RUNG wire#powerrail
      Contact( "Get Sinais de Interlock Falcare".Station[8]."Sinal do job"[6] )
      I_Contact( "BYPASS_MOD_1" )
      I_Contact( "BYPASS_GERAL" )
      I_Contact( "BYPASS_POSTO_60" )
      Coil( "Signals".ProcessInterlock_APLC_Input[1].ModezoneInterlock_APLC_Input[1].StationInterlock_APLC_Input[11].PositionInterlock_APLC_Input[1].EquipmentInterlock_APLC_Input[1].SignalInterlock_APLC_Input[5] )
   END_RUNG
   RUNG wire#powerrail
      Contact( "Get Sinais de Interlock Falcare".Station[8]."Sinal do job"[7] )
      I_Contact( "BYPASS_MOD_1" )
      I_Contact( "BYPASS_GERAL" )
      I_Contact( "BYPASS_POSTO_60" )
      Coil( "Signals".ProcessInterlock_APLC_Input[1].ModezoneInterlock_APLC_Input[1].StationInterlock_APLC_Input[11].PositionInterlock_APLC_Input[1].EquipmentInterlock_APLC_Input[1].SignalInterlock_APLC_Input[6] )
   END_RUNG
   RUNG wire#powerrail
      I_Contact( "Get Sinais de Interlock Falcare".Station[8]."Sinal do job"[9] )
      I_Contact( "BYPASS_MOD_1" )
      I_Contact( "BYPASS_GERAL" )
      I_Contact( "Put Sinais de Interlock Falcare".Bypass_Cortina )
      Coil( "Signals".ProcessInterlock_APLC_Input[1].ModezoneInterlock_APLC_Input[1].StationInterlock_APLC_Input[4].PositionInterlock_APLC_Input[1].EquipmentInterlock_APLC_Input[1].SignalInterlock_APLC_Input[6] )
   END_RUNG
   RUNG wire#powerrail
      I_Contact( "Get Sinais de Interlock Falcare".Station[8]."Sinal do job"[8] )
      I_Contact( "BYPASS_MOD_1" )
      I_Contact( "BYPASS_GERAL" )
      I_Contact( "Put Sinais de Interlock Falcare".Bypass_Cortina )
      Coil( "Signals".ProcessInterlock_APLC_Input[1].ModezoneInterlock_APLC_Input[1].StationInterlock_APLC_Input[4].PositionInterlock_APLC_Input[1].EquipmentInterlock_APLC_Input[1].SignalInterlock_APLC_Input[7] )
   END_RUNG
   RUNG wire#powerrail
      Contact( "AlwaysFALSE" )
      Coil( "Put Sinais de Interlock Falcare".Bypass_Cortina )
   END_RUNG
   // the same network as SCL:
   "Signals".ProcessInterlock_APLC_Input[1].ModezoneInterlock_APLC_Input[1].StationInterlock_APLC_Input[11].PositionInterlock_APLC_Input[1].EquipmentInterlock_APLC_Input[1].SignalInterlock_APLC_Input[1] := "Get Sinais de Interlock Falcare".Station[8]."Sinal do job"[0] AND NOT "BYPASS_MOD_1" AND NOT "BYPASS_GERAL" AND NOT "BYPASS_POSTO_60";
   "Signals".ProcessInterlock_APLC_Input[1].ModezoneInterlock_APLC_Input[1].StationInterlock_APLC_Input[11].PositionInterlock_APLC_Input[1].EquipmentInterlock_APLC_Input[1].SignalInterlock_APLC_Input[2] := "Get Sinais de Interlock Falcare".Station[8]."Sinal do job"[1] AND NOT "BYPASS_MOD_1" AND NOT "BYPASS_GERAL" AND NOT "BYPASS_POSTO_60";
   "Signals".ProcessInterlock_APLC_Input[1].ModezoneInterlock_APLC_Input[1].StationInterlock_APLC_Input[11].PositionInterlock_APLC_Input[1].EquipmentInterlock_APLC_Input[2].SignalInterlock_APLC_Input[2] := NOT "Get Sinais de Interlock Falcare".Station[8]."Sinal do job"[3] AND NOT "BYPASS_MOD_1" AND NOT "BYPASS_GERAL" AND NOT "BYPASS_POSTO_60";
   "Signals".ProcessInterlock_APLC_Input[1].ModezoneInterlock_APLC_Input[1].StationInterlock_APLC_Input[11].PositionInterlock_APLC_Input[1].EquipmentInterlock_APLC_Input[1].SignalInterlock_APLC_Input[3] := "Get Sinais de Interlock Falcare".Station[8]."Sinal do job"[4] AND NOT "BYPASS_MOD_1" AND NOT "BYPASS_GERAL" AND NOT "BYPASS_POSTO_60";
   "Signals".ProcessInterlock_APLC_Input[1].ModezoneInterlock_APLC_Input[1].StationInterlock_APLC_Input[11].PositionInterlock_APLC_Input[1].EquipmentInterlock_APLC_Input[1].SignalInterlock_APLC_Input[4] := "Get Sinais de Interlock Falcare".Station[8]."Sinal do job"[5] AND NOT "BYPASS_MOD_1" AND NOT "BYPASS_GERAL" AND NOT "Get Sinais de Interlock Falcare".Station[8]."Sinal do job"[6] AND NOT "BYPASS_POSTO_60";
   "Signals".ProcessInterlock_APLC_Input[1].ModezoneInterlock_APLC_Input[1].StationInterlock_APLC_Input[11].PositionInterlock_APLC_Input[1].EquipmentInterlock_APLC_Input[1].SignalInterlock_APLC_Input[5] := "Get Sinais de Interlock Falcare".Station[8]."Sinal do job"[6] AND NOT "BYPASS_MOD_1" AND NOT "BYPASS_GERAL" AND NOT "BYPASS_POSTO_60";
   "Signals".ProcessInterlock_APLC_Input[1].ModezoneInterlock_APLC_Input[1].StationInterlock_APLC_Input[11].PositionInterlock_APLC_Input[1].EquipmentInterlock_APLC_Input[1].SignalInterlock_APLC_Input[6] := "Get Sinais de Interlock Falcare".Station[8]."Sinal do job"[7] AND NOT "BYPASS_MOD_1" AND NOT "BYPASS_GERAL" AND NOT "BYPASS_POSTO_60";
   "Signals".ProcessInterlock_APLC_Input[1].ModezoneInterlock_APLC_Input[1].StationInterlock_APLC_Input[4].PositionInterlock_APLC_Input[1].EquipmentInterlock_APLC_Input[1].SignalInterlock_APLC_Input[6] := NOT "Get Sinais de Interlock Falcare".Station[8]."Sinal do job"[9] AND NOT "BYPASS_MOD_1" AND NOT "BYPASS_GERAL" AND NOT "Put Sinais de Interlock Falcare".Bypass_Cortina;
   "Signals".ProcessInterlock_APLC_Input[1].ModezoneInterlock_APLC_Input[1].StationInterlock_APLC_Input[4].PositionInterlock_APLC_Input[1].EquipmentInterlock_APLC_Input[1].SignalInterlock_APLC_Input[7] := NOT "Get Sinais de Interlock Falcare".Station[8]."Sinal do job"[8] AND NOT "BYPASS_MOD_1" AND NOT "BYPASS_GERAL" AND NOT "Put Sinais de Interlock Falcare".Bypass_Cortina;
   "Put Sinais de Interlock Falcare".Bypass_Cortina := "AlwaysFALSE";
END_REGION

REGION Network 13: ALARME IHM TRANSPORTADOR FALCARE
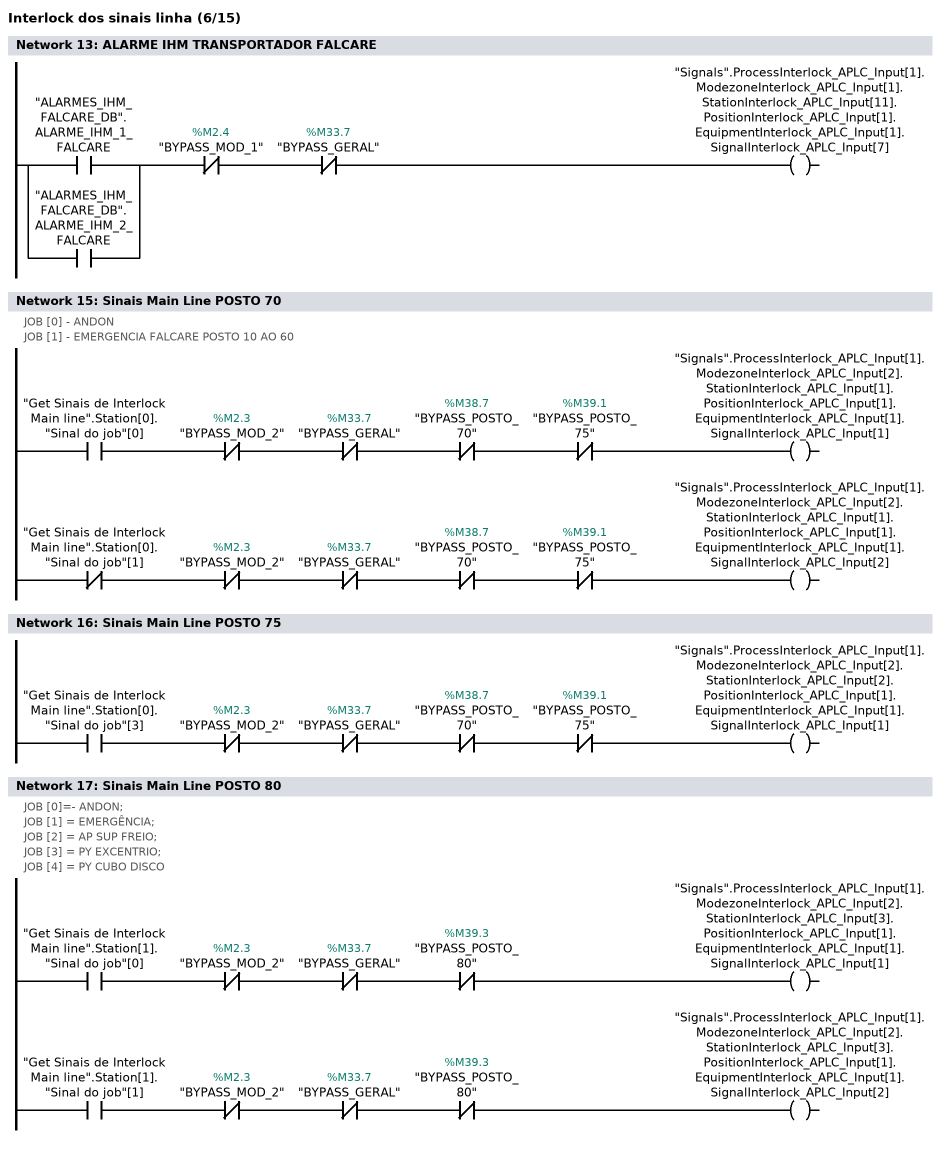
   RUNG wire#powerrail
      Contact( "ALARMES_IHM_FALCARE_DB".ALARME_IHM_1_FALCARE )
      wire#w1
      I_Contact( "BYPASS_MOD_1" )
      I_Contact( "BYPASS_GERAL" )
      Coil( "Signals".ProcessInterlock_APLC_Input[1].ModezoneInterlock_APLC_Input[1].StationInterlock_APLC_Input[11].PositionInterlock_APLC_Input[1].EquipmentInterlock_APLC_Input[1].SignalInterlock_APLC_Input[7] )
   END_RUNG
   RUNG wire#powerrail
      Contact( "ALARMES_IHM_FALCARE_DB".ALARME_IHM_2_FALCARE )
   END_RUNG wire#w1
   // the same network as SCL:
   "Signals".ProcessInterlock_APLC_Input[1].ModezoneInterlock_APLC_Input[1].StationInterlock_APLC_Input[11].PositionInterlock_APLC_Input[1].EquipmentInterlock_APLC_Input[1].SignalInterlock_APLC_Input[7] := ("ALARMES_IHM_FALCARE_DB".ALARME_IHM_1_FALCARE OR "ALARMES_IHM_FALCARE_DB".ALARME_IHM_2_FALCARE) AND NOT "BYPASS_MOD_1" AND NOT "BYPASS_GERAL";
END_REGION

REGION Network 14: Sinais GIRADOR
END_REGION

REGION Network 15: Sinais Main Line POSTO 70
   // JOB [0] - ANDON
   // JOB [1] - EMERGENCIA FALCARE POSTO 10 AO 60
   RUNG wire#powerrail
      Contact( "Get Sinais de Interlock Main line".Station[0]."Sinal do job"[0] )
      I_Contact( "BYPASS_MOD_2" )
      I_Contact( "BYPASS_GERAL" )
      I_Contact( "BYPASS_POSTO_70" )
      I_Contact( "BYPASS_POSTO_75" )
      Coil( "Signals".ProcessInterlock_APLC_Input[1].ModezoneInterlock_APLC_Input[2].StationInterlock_APLC_Input[1].PositionInterlock_APLC_Input[1].EquipmentInterlock_APLC_Input[1].SignalInterlock_APLC_Input[1] )
   END_RUNG
   RUNG wire#powerrail
      I_Contact( "Get Sinais de Interlock Main line".Station[0]."Sinal do job"[1] )
      I_Contact( "BYPASS_MOD_2" )
      I_Contact( "BYPASS_GERAL" )
      I_Contact( "BYPASS_POSTO_70" )
      I_Contact( "BYPASS_POSTO_75" )
      Coil( "Signals".ProcessInterlock_APLC_Input[1].ModezoneInterlock_APLC_Input[2].StationInterlock_APLC_Input[1].PositionInterlock_APLC_Input[1].EquipmentInterlock_APLC_Input[1].SignalInterlock_APLC_Input[2] )
   END_RUNG
   // the same network as SCL:
   "Signals".ProcessInterlock_APLC_Input[1].ModezoneInterlock_APLC_Input[2].StationInterlock_APLC_Input[1].PositionInterlock_APLC_Input[1].EquipmentInterlock_APLC_Input[1].SignalInterlock_APLC_Input[1] := "Get Sinais de Interlock Main line".Station[0]."Sinal do job"[0] AND NOT "BYPASS_MOD_2" AND NOT "BYPASS_GERAL" AND NOT "BYPASS_POSTO_70" AND NOT "BYPASS_POSTO_75";
   "Signals".ProcessInterlock_APLC_Input[1].ModezoneInterlock_APLC_Input[2].StationInterlock_APLC_Input[1].PositionInterlock_APLC_Input[1].EquipmentInterlock_APLC_Input[1].SignalInterlock_APLC_Input[2] := NOT "Get Sinais de Interlock Main line".Station[0]."Sinal do job"[1] AND NOT "BYPASS_MOD_2" AND NOT "BYPASS_GERAL" AND NOT "BYPASS_POSTO_70" AND NOT "BYPASS_POSTO_75";
END_REGION

REGION Network 16: Sinais Main Line POSTO 75
   RUNG wire#powerrail
      Contact( "Get Sinais de Interlock Main line".Station[0]."Sinal do job"[3] )
      I_Contact( "BYPASS_MOD_2" )
      I_Contact( "BYPASS_GERAL" )
      I_Contact( "BYPASS_POSTO_70" )
      I_Contact( "BYPASS_POSTO_75" )
      Coil( "Signals".ProcessInterlock_APLC_Input[1].ModezoneInterlock_APLC_Input[2].StationInterlock_APLC_Input[2].PositionInterlock_APLC_Input[1].EquipmentInterlock_APLC_Input[1].SignalInterlock_APLC_Input[1] )
   END_RUNG
   // the same network as SCL:
   "Signals".ProcessInterlock_APLC_Input[1].ModezoneInterlock_APLC_Input[2].StationInterlock_APLC_Input[2].PositionInterlock_APLC_Input[1].EquipmentInterlock_APLC_Input[1].SignalInterlock_APLC_Input[1] := "Get Sinais de Interlock Main line".Station[0]."Sinal do job"[3] AND NOT "BYPASS_MOD_2" AND NOT "BYPASS_GERAL" AND NOT "BYPASS_POSTO_70" AND NOT "BYPASS_POSTO_75";
END_REGION

